  MoveL 5119 to (-200, -30.3, 0.2) mm, rotated rx 1.14 ry 0 rz 180 deg; joints [20.999, -64.73, 124.107, -155.961, 61.604, 79.168]
  MoveL 5120 to (0, -30.3, 0.2) mm, rotated rx 1.14 ry 0 rz 180 deg; joints [18.154, -55.53, 108.18, -157.586, 54.796, 77.769]
  MoveL 5121 to (0, -29.7, 0.2) mm, rotated rx 0 ry 0 rz 180 deg; joints [18.189, -55.157, 108.238, -157.658, 55.202, 76.801]
  MoveL 5122 to (-200, -29.7, 0.2) mm, rotated rx 0 ry 0 rz 180 deg; joints [21.039, -64.279, 124.171, -156.029, 62.083, 78.241]
  MoveL 5123 to (-200, -29.1, 0.2) mm, rotated rx 0 ry 0 rz 180 deg; joints [21.039, -64.245, 124.178, -156.038, 62.121, 78.259]
  MoveL 5124 to (0, -29.1, 0.2) mm, rotated rx 0 ry 0 rz 180 deg; joints [18.189, -55.13, 108.244, -157.667, 55.234, 76.816]
  MoveL 5125 to (0, -28.5, 0.2) mm, rotated rx 0 ry 0 rz 180 deg; joints [18.189, -55.102, 108.25, -157.676, 55.266, 76.832]
  MoveL 5126 to (-200, -28.5, 0.2) mm, rotated rx 0 ry 0 rz 180 deg; joints [21.039, -64.211, 124.185, -156.046, 62.158, 78.278]
  MoveL 5127 to (-200, -27.9, 0.2) mm, rotated rx 0 ry 0 rz 180 deg; joints [21.039, -64.177, 124.192, -156.055, 62.195, 78.297]
  MoveL 5128 to (0, -27.9, 0.2) mm, rotated rx 0 ry 0 rz 180 deg; joints [18.189, -55.074, 108.257, -157.685, 55.297, 76.848]
  MoveL 5129 to (0, -27.3, 0.2) mm, rotated rx 0 ry 0 rz 180 deg; joints [18.189, -55.046, 108.263, -157.694, 55.329, 76.864]
  MoveL 5130 to (-200, -27.3, 0.2) mm, rotated rx 0 ry 0 rz 180 deg; joints [21.039, -64.143, 124.198, -156.064, 62.232, 78.316]
  MoveL 5131 to (-200, -26.7, 0.2) mm, rotated rx 0 ry 0 rz 180 deg; joints [21.039, -64.109, 124.205, -156.072, 62.269, 78.334]
  MoveL 5132 to (0, -26.7, 0.2) mm, rotated rx 0 ry 0 rz 180 deg; joints [18.189, -55.018, 108.269, -157.703, 55.361, 76.88]
  MoveL 5133 to (0, -26.1, 0.2) mm, rotated rx 0 ry 0 rz 180 deg; joints [18.189, -54.99, 108.275, -157.712, 55.392, 76.895]
  MoveL 5134 to (-200, -26.1, 0.2) mm, rotated rx 0 ry 0 rz 180 deg; joints [21.039, -64.075, 124.212, -156.081, 62.307, 78.353]
  MoveL 5135 to (-200, -25.5, 0.2) mm, rotated rx 0 ry 0 rz 180 deg; joints [21.039, -64.041, 124.218, -156.09, 62.344, 78.372]
  MoveL 5136 to (0, -25.5, 0.2) mm, rotated rx 0 ry 0 rz 180 deg; joints [18.189, -54.962, 108.281, -157.721, 55.424, 76.911]
  MoveL 5137 to (0, -24.9, 0.2) mm, rotated rx 0 ry 0 rz 180 deg; joints [18.189, -54.934, 108.288, -157.73, 55.455, 76.927]
  MoveL 5138 to (-200, -24.9, 0.2) mm, rotated rx 0 ry 0 rz 180 deg; joints [21.039, -64.007, 124.225, -156.098, 62.381, 78.39]
  MoveL 5139 to (-200, -24.3, 0.2) mm, rotated rx 0 ry 0 rz 180 deg; joints [21.039, -63.973, 124.232, -156.107, 62.418, 78.409]
  MoveL 5140 to (0, -24.3, 0.2) mm, rotated rx 0 ry 0 rz 180 deg; joints [18.189, -54.906, 108.294, -157.739, 55.487, 76.942]
  MoveL 5141 to (0, -23.7, 0.2) mm, rotated rx 0 ry 0 rz 180 deg; joints [18.189, -54.878, 108.3, -157.748, 55.519, 76.958]
  MoveL 5142 to (-200, -23.7, 0.2) mm, rotated rx 0 ry 0 rz 180 deg; joints [21.039, -63.939, 124.238, -156.116, 62.455, 78.427]
  MoveL 5143 to (-200, -23.1, 0.2) mm, rotated rx 0 ry 0 rz 180 deg; joints [21.039, -63.905, 124.245, -156.124, 62.493, 78.446]
  MoveL 5144 to (0, -23.1, 0.2) mm, rotated rx 0 ry 0 rz 180 deg; joints [18.189, -54.849, 108.306, -157.757, 55.55, 76.974]
  MoveL 5145 to (0, -22.5, 0.2) mm, rotated rx 0 ry 0 rz 180 deg; joints [18.189, -54.821, 108.312, -157.766, 55.582, 76.989]
  MoveL 5146 to (-200, -22.5, 0.2) mm, rotated rx 0 ry 0 rz 180 deg; joints [21.039, -63.871, 124.251, -156.133, 62.53, 78.464]
  MoveL 5147 to (-200, -21.9, 0.2) mm, rotated rx 0 ry 0 rz 180 deg; joints [21.039, -63.836, 124.258, -156.141, 62.567, 78.483]
  MoveL 5148 to (0, -21.9, 0.2) mm, rotated rx 0 ry 0 rz 180 deg; joints [18.189, -54.793, 108.318, -157.775, 55.613, 77.005]
  MoveL 5149 to (0, -21.3, 0.2) mm, rotated rx 0 ry 0 rz 180 deg; joints [18.189, -54.765, 108.324, -157.783, 55.645, 77.021]
  MoveL 5150 to (-200, -21.3, 0.2) mm, rotated rx 0 ry 0 rz 180 deg; joints [21.039, -63.802, 124.264, -156.15, 62.604, 78.501]
  MoveL 5151 to (-200, -20.7, 0.2) mm, rotated rx 0 ry 0 rz 180 deg; joints [21.039, -63.768, 124.271, -156.158, 62.641, 78.52]
  MoveL 5152 to (0, -20.7, 0.2) mm, rotated rx 0 ry 0 rz 180 deg; joints [18.189, -54.737, 108.33, -157.792, 55.676, 77.036]
  MoveL 5153 to (0, -20.1, 0.2) mm, rotated rx 0 ry 0 rz 180 deg; joints [18.189, -54.709, 108.335, -157.801, 55.708, 77.052]
  MoveL 5154 to (-200, -20.1, 0.2) mm, rotated rx 0 ry 0 rz 180 deg; joints [21.039, -63.734, 124.277, -156.167, 62.678, 78.538]
  MoveL 5155 to (-200, -19.5, 0.2) mm, rotated rx 0 ry 0 rz 180 deg; joints [21.039, -63.7, 124.283, -156.175, 62.716, 78.557]
  MoveL 5156 to (0, -19.5, 0.2) mm, rotated rx 0 ry 0 rz 180 deg; joints [18.189, -54.681, 108.341, -157.81, 55.739, 77.067]
  MoveL 5157 to (0, -18.9, 0.2) mm, rotated rx 0 ry 0 rz 180 deg; joints [18.189, -54.652, 108.347, -157.818, 55.771, 77.083]
  MoveL 5158 to (-200, -18.9, 0.2) mm, rotated rx 0 ry 0 rz 180 deg; joints [21.039, -63.665, 124.29, -156.184, 62.753, 78.575]
  MoveL 5159 to (-200, -18.3, 0.2) mm, rotated rx 0 ry 0 rz 180 deg; joints [21.039, -63.631, 124.296, -156.192, 62.79, 78.594]
  MoveL 5160 to (0, -18.3, 0.2) mm, rotated rx 0 ry 0 rz 180 deg; joints [18.189, -54.624, 108.353, -157.827, 55.802, 77.099]
  MoveL 5161 to (0, -17.7, 0.2) mm, rotated rx 0 ry 0 rz 180 deg; joints [18.189, -54.596, 108.359, -157.836, 55.834, 77.114]
  MoveL 5162 to (-200, -17.7, 0.2) mm, rotated rx 0 ry 0 rz 180 deg; joints [21.039, -63.597, 124.302, -156.201, 62.827, 78.612]
  MoveL 5163 to (-200, -17.1, 0.2) mm, rotated rx 0 ry 0 rz 180 deg; joints [21.039, -63.562, 124.308, -156.209, 62.864, 78.631]
  MoveL 5164 to (0, -17.1, 0.2) mm, rotated rx 0 ry 0 rz 180 deg; joints [18.189, -54.568, 108.364, -157.845, 55.865, 77.13]
  MoveL 5165 to (0, -16.5, 0.2) mm, rotated rx 0 ry 0 rz 180 deg; joints [18.189, -54.539, 108.37, -157.853, 55.897, 77.145]
  MoveL 5166 to (-200, -16.5, 0.2) mm, rotated rx 0 ry 0 rz 180 deg; joints [21.039, -63.528, 124.315, -156.217, 62.901, 78.649]
  MoveL 5167 to (-200, -15.9, 0.2) mm, rotated rx 0 ry 0 rz 180 deg; joints [21.039, -63.494, 124.321, -156.226, 62.938, 78.667]
  MoveL 5168 to (0, -15.9, 0.2) mm, rotated rx 0 ry 0 rz 180 deg; joints [18.189, -54.511, 108.376, -157.862, 55.928, 77.161]
  MoveL 5169 to (0, -15.3, 0.2) mm, rotated rx 0 ry 0 rz 180 deg; joints [18.189, -54.483, 108.381, -157.871, 55.96, 77.176]
  MoveL 5170 to (-200, -15.3, 0.2) mm, rotated rx 0 ry 0 rz 180 deg; joints [21.039, -63.459, 124.327, -156.234, 62.975, 78.686]
  MoveL 5171 to (-200, -14.7, 0.2) mm, rotated rx 0 ry 0 rz 180 deg; joints [21.039, -63.425, 124.333, -156.242, 63.012, 78.704]
  MoveL 5172 to (0, -14.7, 0.2) mm, rotated rx 0 ry 0 rz 180 deg; joints [18.189, -54.454, 108.387, -157.879, 55.991, 77.191]
  MoveL 5173 to (0, -14.1, 0.2) mm, rotated rx 0 ry 0 rz 180 deg; joints [18.189, -54.426, 108.393, -157.888, 56.023, 77.207]
  MoveL 5174 to (-200, -14.1, 0.2) mm, rotated rx 0 ry 0 rz 180 deg; joints [21.039, -63.39, 124.339, -156.251, 63.049, 78.722]
  MoveL 5175 to (-200, -13.5, 0.2) mm, rotated rx 0 ry 0 rz 180 deg; joints [21.039, -63.356, 124.345, -156.259, 63.087, 78.741]
  MoveL 5176 to (0, -13.5, 0.2) mm, rotated rx 0 ry 0 rz 180 deg; joints [18.189, -54.398, 108.398, -157.896, 56.054, 77.222]
  MoveL 5177 to (0, -12.9, 0.2) mm, rotated rx 0 ry 0 rz 180 deg; joints [18.189, -54.369, 108.404, -157.905, 56.086, 77.238]
  MoveL 5178 to (-200, -12.9, 0.2) mm, rotated rx 0 ry 0 rz 180 deg; joints [21.039, -63.321, 124.351, -156.267, 63.124, 78.759]
  MoveL 5179 to (-200, -12.3, 0.2) mm, rotated rx 0 ry 0 rz 180 deg; joints [21.039, -63.287, 124.357, -156.275, 63.161, 78.777]
  MoveL 5180 to (0, -12.3, 0.2) mm, rotated rx 0 ry 0 rz 180 deg; joints [18.189, -54.341, 108.409, -157.914, 56.117, 77.253]
  MoveL 5181 to (0, -11.7, 0.2) mm, rotated rx 0 ry 0 rz 180 deg; joints [18.189, -54.312, 108.415, -157.922, 56.148, 77.268]
  MoveL 5182 to (-200, -11.7, 0.2) mm, rotated rx 0 ry 0 rz 180 deg; joints [21.039, -63.252, 124.363, -156.284, 63.198, 78.795]
  MoveL 5183 to (-200, -11.1, 0.2) mm, rotated rx 0 ry 0 rz 180 deg; joints [21.039, -63.218, 124.369, -156.292, 63.235, 78.814]
  MoveL 5184 to (0, -11.1, 0.2) mm, rotated rx 0 ry 0 rz 180 deg; joints [18.189, -54.284, 108.42, -157.931, 56.18, 77.284]
  MoveL 5185 to (0, -10.5, 0.2) mm, rotated rx 0 ry 0 rz 180 deg; joints [18.189, -54.256, 108.426, -157.939, 56.211, 77.299]
  MoveL 5186 to (-200, -10.5, 0.2) mm, rotated rx 0 ry 0 rz 180 deg; joints [21.039, -63.183, 124.375, -156.3, 63.272, 78.832]
  MoveL 5187 to (-200, -9.9, 0.2) mm, rotated rx 0 ry 0 rz 180 deg; joints [21.039, -63.149, 124.381, -156.308, 63.309, 78.85]
  MoveL 5188 to (0, -9.9, 0.2) mm, rotated rx 0 ry 0 rz 180 deg; joints [18.189, -54.227, 108.431, -157.948, 56.243, 77.314]
  MoveL 5189 to (0, -9.3, 0.2) mm, rotated rx 0 ry 0 rz 180 deg; joints [18.189, -54.199, 108.436, -157.956, 56.274, 77.33]
  MoveL 5190 to (-200, -9.3, 0.2) mm, rotated rx 0 ry 0 rz 180 deg; joints [21.039, -63.114, 124.387, -156.316, 63.346, 78.868]
  MoveL 5191 to (-200, -8.7, 0.2) mm, rotated rx 0 ry 0 rz 180 deg; joints [21.039, -63.079, 124.392, -156.325, 63.383, 78.886]
  MoveL 5192 to (0, -8.7, 0.2) mm, rotated rx 0 ry 0 rz 180 deg; joints [18.189, -54.17, 108.442, -157.965, 56.305, 77.345]
  MoveL 5193 to (0, -8.1, 0.2) mm, rotated rx 0 ry 0 rz 180 deg; joints [18.189, -54.141, 108.447, -157.973, 56.337, 77.36]
  MoveL 5194 to (-200, -8.1, 0.2) mm, rotated rx 0 ry 0 rz 180 deg; joints [21.039, -63.045, 124.398, -156.333, 63.42, 78.904]
  MoveL 5195 to (-200, -7.5, 0.2) mm, rotated rx 0 ry 0 rz 180 deg; joints [21.039, -63.01, 124.404, -156.341, 63.457, 78.923]
  MoveL 5196 to (0, -7.5, 0.2) mm, rotated rx 0 ry 0 rz 180 deg; joints [18.189, -54.113, 108.452, -157.982, 56.368, 77.375]
  MoveL 5197 to (0, -6.9, 0.2) mm, rotated rx 0 ry 0 rz 180 deg; joints [18.189, -54.084, 108.457, -157.99, 56.399, 77.391]
  MoveL 5198 to (-200, -6.9, 0.2) mm, rotated rx 0 ry 0 rz 180 deg; joints [21.039, -62.975, 124.409, -156.349, 63.494, 78.941]
  MoveL 5199 to (-200, -6.3, 0.2) mm, rotated rx 0 ry 0 rz 180 deg; joints [21.039, -62.941, 124.415, -156.357, 63.531, 78.959]
  MoveL 5200 to (0, -6.3, 0.2) mm, rotated rx 0 ry 0 rz 180 deg; joints [18.189, -54.056, 108.463, -157.998, 56.431, 77.406]
  MoveL 5201 to (0, -5.7, 0.2) mm, rotated rx 0 ry 0 rz 180 deg; joints [18.189, -54.027, 108.468, -158.007, 56.462, 77.421]
  MoveL 5202 to (-200, -5.7, 0.2) mm, rotated rx 0 ry 0 rz 180 deg; joints [21.039, -62.906, 124.421, -156.365, 63.568, 78.977]
  MoveL 5203 to (-200, -5.1, 0.2) mm, rotated rx 0 ry 0 rz 180 deg; joints [21.039, -62.871, 124.426, -156.373, 63.605, 78.995]
  MoveL 5204 to (0, -5.1, 0.2) mm, rotated rx 0 ry 0 rz 180 deg; joints [18.189, -53.999, 108.473, -158.015, 56.493, 77.436]
  MoveL 5205 to (0, -4.5, 0.2) mm, rotated rx 0 ry 0 rz 180 deg; joints [18.189, -53.97, 108.478, -158.024, 56.525, 77.451]
  MoveL 5206 to (-200, -4.5, 0.2) mm, rotated rx 0 ry 0 rz 180 deg; joints [21.039, -62.836, 124.432, -156.381, 63.642, 79.013]
  MoveL 5207 to (-200, -3.9, 0.2) mm, rotated rx 0 ry 0 rz 180 deg; joints [21.039, -62.802, 124.437, -156.389, 63.679, 79.031]
  MoveL 5208 to (0, -3.9, 0.2) mm, rotated rx 0 ry 0 rz 180 deg; joints [18.189, -53.941, 108.483, -158.032, 56.556, 77.466]
  MoveL 5209 to (0, -3.3, 0.2) mm, rotated rx 0 ry 0 rz 180 deg; joints [18.189, -53.913, 108.488, -158.04, 56.587, 77.481]
  MoveL 5210 to (-200, -3.3, 0.2) mm, rotated rx 0 ry 0 rz 180 deg; joints [21.039, -62.767, 124.443, -156.397, 63.716, 79.049]
  MoveL 5211 to (-200, -2.7, 0.2) mm, rotated rx 0 ry 0 rz 180 deg; joints [21.039, -62.732, 124.448, -156.405, 63.753, 79.067]
  MoveL 5212 to (0, -2.7, 0.2) mm, rotated rx 0 ry 0 rz 180 deg; joints [18.189, -53.884, 108.493, -158.049, 56.619, 77.497]
  MoveL 5213 to (0, -2.1, 0.2) mm, rotated rx 0 ry 0 rz 180 deg; joints [18.189, -53.855, 108.498, -158.057, 56.65, 77.512]
  MoveL 5214 to (-200, -2.1, 0.2) mm, rotated rx 0 ry 0 rz 180 deg; joints [21.039, -62.697, 124.454, -156.413, 63.789, 79.085]
  MoveL 5215 to (-200, -1.5, 0.2) mm, rotated rx 0 ry 0 rz 180 deg; joints [21.039, -62.662, 124.459, -156.421, 63.826, 79.103]
  MoveL 5216 to (0, -1.5, 0.2) mm, rotated rx 0 ry 0 rz 180 deg; joints [18.189, -53.826, 108.503, -158.065, 56.681, 77.527]
  MoveL 5217 to (0, -0.9, 0.2) mm, rotated rx 0 ry 0 rz 180 deg; joints [18.189, -53.798, 108.508, -158.073, 56.712, 77.542]
  MoveL 5218 to (-200, -0.9, 0.2) mm, rotated rx 0 ry 0 rz 180 deg; joints [21.039, -62.627, 124.465, -156.429, 63.863, 79.121]
  MoveL 5219 to (-200, -0.3, 0.2) mm, rotated rx 0 ry 0 rz 180 deg; joints [21.039, -62.592, 124.47, -156.437, 63.9, 79.139]
  MoveL 5220 to (0, -0.3, 0.2) mm, rotated rx 0 ry 0 rz 180 deg; joints [18.189, -53.769, 108.513, -158.082, 56.744, 77.557]
  MoveL 5221 to (0, 0, 0.2) mm, rotated rx 0 ry 0 rz 180 deg; joints [18.189, -53.755, 108.515, -158.086, 56.759, 77.564]
  MoveL 5222 to (-200, 0, 0.2) mm, rotated rx 0 ry 0 rz 180 deg; joints [21.039, -62.575, 124.473, -156.44, 63.918, 79.148]
  Sollgeschwindigkeit (200.0 mm/s)
  MoveL 5223 to (-200, 0, -44.8) mm, rotated rx 0 ry 0 rz 180 deg; joints [22.93, -61.804, 123.11, -154.254, 63.757, 77.962]
  END

--- program CBL1 (robot KUKA KR 30 HA) ---
  Glatt(1)
  Sollgeschwindigkeit (1000.0 mm/s)
  Referenz erstellen.: Reference SW
  Werkzeug setzen: PlasticPos800
  Anzeigen PlasticPos800
  MoveJ 1 to (-41.72, -40.46, 48.98) mm, rotated rx 90 ry 0 rz 90 deg; joints [0.027, -82.593, 139.4, -179.968, 56.807, 179.983]
  MoveL 2 to (-41.72, -40.46, 48.98) mm, rotated rx 90 ry 0 rz 90 deg; joints [0.027, -82.593, 139.4, -179.968, 56.807, 179.983]
  MoveL 3 to (-41.72, -40.46, 48.98) mm, rotated rx 90 ry 0 rz 90 deg; joints [0.027, -82.593, 139.4, -179.968, 56.807, 179.983]
  MoveL 4 to (-41.72, -40.46, 48.98) mm, rotated rx 90 ry 0 rz 90 deg; joints [0.027, -82.593, 139.4, -179.968, 56.807, 179.983]
  Sollgeschwindigkeit (50.0 mm/s)
  MoveL 5 to (-32.85, -40.57, 48.4) mm, rotated rx 90 ry 0 rz 90 deg; joints [0.058, -82.072, 138.764, -179.93, 56.692, 179.962]
  MoveL 6 to (-23.97, -40.69, 47.75) mm, rotated rx 90 ry 0 rz 90 deg; joints [0.094, -81.555, 138.126, -179.887, 56.571, 179.938]
  MoveL 7 to (-15.09, -40.74, 47.81) mm, rotated rx 90 ry 0 rz 90 deg; joints [0.089, -81.036, 137.485, -179.893, 56.449, 179.941]
  MoveL 8 to (-6.28, -40.47, 49.1) mm, rotated rx 90 ry 0 rz 90 deg; joints [0.02, -80.506, 136.856, -179.976, 56.35, 179.987]
  MoveL 9 to (-0.84, -39.84, 50.5) mm, rotated rx 90 ry 0 rz 90 deg; joints [-0.055, -80.152, 136.477, -180.066, 56.326, 180.037]
  MoveL 10 to (4.48, -38.76, 52.1) mm, rotated rx 90 ry 0 rz 90 deg; joints [-0.14, -79.779, 136.116, -180.168, 56.337, 180.093]
  MoveL 11 to (9.75, -37.21, 53.58) mm, rotated rx 90 ry 0 rz 90 deg; joints [-0.218, -79.383, 135.768, -180.262, 56.385, 180.145]
  MoveL 12 to (14.99, -35.35, 54.76) mm, rotated rx 90 ry 0 rz 90 deg; joints [-0.279, -78.971, 135.428, -180.335, 56.457, 180.185]
  MoveL 13 to (20.23, -33.45, 55.56) mm, rotated rx 90 ry 0 rz 90 deg; joints [-0.32, -78.559, 135.087, -180.383, 56.528, 180.212]
  MoveL 14 to (25.53, -31.86, 55.96) mm, rotated rx 90 ry 0 rz 90 deg; joints [-0.339, -78.165, 134.733, -180.407, 56.569, 180.224]
  MoveL 15 to (31.11, -31.04, 56.06) mm, rotated rx 90 ry 0 rz 90 deg; joints [-0.343, -77.802, 134.34, -180.411, 56.539, 180.227]
  MoveL 16 to (37.22, -31.47, 56) mm, rotated rx 90 ry 0 rz 90 deg; joints [-0.338, -77.485, 133.88, -180.405, 56.395, 180.224]
  MoveL 17 to (43.65, -32.9, 55.86) mm, rotated rx 90 ry 0 rz 90 deg; joints [-0.329, -77.209, 133.372, -180.396, 56.164, 180.22]
  MoveL 18 to (50.35, -33.59, 55.79) mm, rotated rx 90 ry 0 rz 90 deg; joints [-0.323, -76.875, 132.859, -180.39, 55.985, 180.218]
  MoveL 19 to (57.02, -32.75, 55.87) mm, rotated rx 90 ry 0 rz 90 deg; joints [-0.325, -76.455, 132.381, -180.393, 55.926, 180.22]
  MoveL 20 to (63.44, -31.36, 56.01) mm, rotated rx 90 ry 0 rz 90 deg; joints [-0.33, -76.02, 131.931, -180.399, 55.912, 180.224]
  MoveL 21 to (69.49, -31.08, 56.06) mm, rotated rx 90 ry 0 rz 90 deg; joints [-0.331, -75.67, 131.484, -180.401, 55.815, 180.225]
  MoveL 22 to (75.02, -32, 55.94) mm, rotated rx 90 ry 0 rz 90 deg; joints [-0.323, -75.417, 131.048, -180.392, 55.631, 180.221]
  MoveL 23 to (80.31, -33.64, 55.49) mm, rotated rx 90 ry 0 rz 90 deg; joints [-0.3, -75.218, 130.615, -180.364, 55.397, 180.207]
  MoveL 24 to (85.55, -35.55, 54.65) mm, rotated rx 90 ry 0 rz 90 deg; joints [-0.257, -75.036, 130.178, -180.313, 55.143, 180.179]
  MoveL 25 to (93.19, -38.13, 52.78) mm, rotated rx 90 ry 0 rz 90 deg; joints [-0.163, -74.758, 129.545, -180.2, 54.787, 180.115]
  MoveL 26 to (100.91, -39.85, 50.48) mm, rotated rx 90 ry 0 rz 90 deg; joints [-0.049, -74.427, 128.922, -180.061, 54.495, 180.035]
  MoveL 27 to (108.88, -40.62, 48.59) mm, rotated rx 90 ry 0 rz 90 deg; joints [0.042, -74.031, 128.298, -179.948, 54.266, 179.969]
  MoveL 28 to (117.07, -40.74, 47.7) mm, rotated rx 90 ry 0 rz 90 deg; joints [0.085, -73.589, 127.669, -179.895, 54.08, 179.938]
  MoveL 29 to (125.29, -40.67, 47.82) mm, rotated rx 90 ry 0 rz 90 deg; joints [0.079, -73.136, 127.039, -179.903, 53.902, 179.943]
  MoveL 30 to (133.51, -40.57, 48.46) mm, rotated rx 90 ry 0 rz 90 deg; joints [0.048, -72.683, 126.408, -179.941, 53.724, 179.965]
  MoveL 31 to (141.72, -40.46, 48.98) mm, rotated rx 90 ry 0 rz 90 deg; joints [0.023, -72.231, 125.774, -179.972, 53.543, 179.983]
  Sollgeschwindigkeit (1000.0 mm/s)
  MoveL 32 to (141.72, -40.46, 48.98) mm, rotated rx 90 ry 0 rz 90 deg; joints [0.023, -72.231, 125.774, -179.972, 53.543, 179.983]
  MoveL 33 to (141.72, -40.46, 48.98) mm, rotated rx 90 ry 0 rz 90 deg; joints [0.023, -72.231, 125.774, -179.972, 53.543, 179.983]
  Sollgeschwindigkeit (1000.0 mm/s)
  MoveL 34 to (145.1, -41.25, 44.7) mm, rotated rx 90 ry 0 rz 90 deg; joints [0.224, -72.088, 125.494, -179.721, 53.406, 179.834]
  MoveL 35 to (145.1, -41.25, 44.7) mm, rotated rx 90 ry 0 rz 90 deg; joints [0.224, -72.088, 125.494, -179.721, 53.406, 179.834]
  MoveL 36 to (145.1, -41.25, 44.7) mm, rotated rx 90 ry 0 rz 90 deg; joints [0.224, -72.088, 125.494, -179.721, 53.406, 179.834]
  Sollgeschwindigkeit (50.0 mm/s)
  MoveL 37 to (141.7, -41.25, 42.87) mm, rotated rx 90 ry 0 rz 90 deg; joints [0.312, -72.273, 125.758, -179.612, 53.486, 179.769]
  MoveL 38 to (137.92, -41.25, 41.96) mm, rotated rx 90 ry 0 rz 90 deg; joints [0.355, -72.478, 126.05, -179.558, 53.573, 179.738]
  MoveL 39 to (134, -41.25, 41.48) mm, rotated rx 90 ry 0 rz 90 deg; joints [0.379, -72.691, 126.353, -179.529, 53.663, 179.721]
  MoveL 40 to (130.09, -41.25, 41.08) mm, rotated rx 90 ry 0 rz 90 deg; joints [0.4, -72.903, 126.655, -179.505, 53.752, 179.707]
  MoveL 41 to (126.21, -41.24, 40.71) mm, rotated rx 90 ry 0 rz 90 deg; joints [0.419, -73.115, 126.954, -179.481, 53.84, 179.694]
  MoveL 42 to (118.64, -41.24, 39.88) mm, rotated rx 90 ry 0 rz 90 deg; joints [0.461, -73.528, 127.535, -179.43, 54.008, 179.665]
  MoveL 43 to (111.13, -41.25, 38.67) mm, rotated rx 90 ry 0 rz 90 deg; joints [0.523, -73.939, 128.109, -179.355, 54.171, 179.623]
  MoveL 44 to (104.5, -41.27, 37.04) mm, rotated rx 90 ry 0 rz 90 deg; joints [0.605, -74.303, 128.613, -179.255, 54.312, 179.565]
  MoveL 45 to (98.04, -41.26, 34.74) mm, rotated rx 90 ry 0 rz 90 deg; joints [0.721, -74.656, 129.102, -179.113, 54.449, 179.485]
  MoveL 46 to (91.88, -41.2, 31.62) mm, rotated rx 90 ry 0 rz 90 deg; joints [0.879, -74.99, 129.567, -178.922, 54.581, 179.375]
  MoveL 47 to (86.28, -41.2, 27.66) mm, rotated rx 90 ry 0 rz 90 deg; joints [1.079, -75.296, 129.985, -178.678, 54.697, 179.236]
  MoveL 48 to (80.96, -41.38, 22.17) mm, rotated rx 90 ry 0 rz 90 deg; joints [1.356, -75.594, 130.373, -178.34, 54.791, 179.043]
  MoveL 49 to (76.3, -41.22, 15.86) mm, rotated rx 90 ry 0 rz 90 deg; joints [1.677, -75.835, 130.715, -177.95, 54.897, 178.821]
  MoveL 50 to (73.92, -40.67, 12.58) mm, rotated rx 90 ry 0 rz 90 deg; joints [1.844, -75.931, 130.898, -177.748, 54.988, 178.708]
  MoveL 51 to (71.58, -39.57, 9.53) mm, rotated rx 90 ry 0 rz 90 deg; joints [2.001, -75.994, 131.09, -177.561, 55.121, 178.605]
  MoveL 52 to (69.42, -37.75, 7.01) mm, rotated rx 90 ry 0 rz 90 deg; joints [2.131, -76.007, 131.286, -177.408, 55.306, 178.524]
  MoveL 53 to (67.55, -35.05, 5.3) mm, rotated rx 90 ry 0 rz 90 deg; joints [2.22, -75.955, 131.48, -177.307, 55.555, 178.476]
  MoveL 54 to (65.46, -30.42, 4.14) mm, rotated rx 90 ry 0 rz 90 deg; joints [2.283, -75.806, 131.734, -177.245, 55.959, 178.457]
  MoveL 55 to (63.59, -25.34, 3.78) mm, rotated rx 90 ry 0 rz 90 deg; joints [2.305, -75.618, 131.981, -177.233, 56.394, 178.468]
  MoveL 56 to (61.65, -20.55, 3.71) mm, rotated rx 90 ry 0 rz 90 deg; joints [2.312, -75.447, 132.227, -177.237, 56.81, 178.487]
  MoveL 57 to (59.77, -17.22, 3.72) mm, rotated rx 90 ry 0 rz 90 deg; joints [2.315, -75.355, 132.436, -177.243, 57.111, 178.502]
  MoveL 58 to (57.13, -13.98, 3.77) mm, rotated rx 90 ry 0 rz 90 deg; joints [2.318, -75.309, 132.7, -177.248, 57.421, 178.518]
  MoveL 59 to (55.51, -12.44, 3.79) mm, rotated rx 90 ry 0 rz 90 deg; joints [2.32, -75.305, 132.851, -177.251, 57.576, 178.525]
  MoveL 60 to (53.83, -11.08, 3.81) mm, rotated rx 90 ry 0 rz 90 deg; joints [2.323, -75.316, 133.004, -177.252, 57.718, 178.531]
  MoveL 61 to (52.14, -9.99, 3.81) mm, rotated rx 90 ry 0 rz 90 deg; joints [2.327, -75.342, 133.153, -177.251, 57.84, 178.536]
  MoveL 62 to (50, -9.51, 3.8) mm, rotated rx 90 ry 0 rz 90 deg; joints [2.331, -75.43, 133.322, -177.248, 57.923, 178.538]
  MoveL 63 to (47.86, -9.99, 3.81) mm, rotated rx 90 ry 0 rz 90 deg; joints [2.336, -75.574, 133.473, -177.243, 57.929, 178.536]
  MoveL 64 to (46.17, -11.08, 3.81) mm, rotated rx 90 ry 0 rz 90 deg; joints [2.339, -75.731, 133.577, -177.238, 57.876, 178.53]
  MoveL 65 to (44.49, -12.44, 3.79) mm, rotated rx 90 ry 0 rz 90 deg; joints [2.343, -75.904, 133.675, -177.23, 57.801, 178.523]
  MoveL 66 to (42.87, -13.98, 3.77) mm, rotated rx 90 ry 0 rz 90 deg; joints [2.348, -76.084, 133.764, -177.222, 57.711, 178.515]
  MoveL 67 to (40.23, -17.22, 3.72) mm, rotated rx 90 ry 0 rz 90 deg; joints [2.356, -76.422, 133.894, -177.207, 57.503, 178.498]
  MoveL 68 to (38.35, -20.55, 3.71) mm, rotated rx 90 ry 0 rz 90 deg; joints [2.36, -76.725, 133.963, -177.194, 57.27, 178.482]
  MoveL 69 to (36.41, -25.34, 3.78) mm, rotated rx 90 ry 0 rz 90 deg; joints [2.361, -77.117, 134.005, -177.182, 56.92, 178.461]
  MoveL 70 to (34.54, -30.42, 4.14) mm, rotated rx 90 ry 0 rz 90 deg; joints [2.346, -77.522, 134.034, -177.187, 56.543, 178.448]
  MoveL 71 to (32.45, -35.05, 5.3) mm, rotated rx 90 ry 0 rz 90 deg; joints [2.291, -77.915, 134.089, -177.243, 56.205, 178.466]
  MoveL 72 to (30.58, -37.75, 7.01) mm, rotated rx 90 ry 0 rz 90 deg; joints [2.206, -78.182, 134.17, -177.339, 56.016, 178.512]
  MoveL 73 to (28.42, -39.57, 9.53) mm, rotated rx 90 ry 0 rz 90 deg; joints [2.079, -78.417, 134.294, -177.489, 55.902, 178.592]
  MoveL 74 to (26.08, -40.67, 12.58) mm, rotated rx 90 ry 0 rz 90 deg; joints [1.925, -78.62, 134.448, -177.674, 55.85, 178.694]
  MoveL 75 to (23.7, -41.22, 15.86) mm, rotated rx 90 ry 0 rz 90 deg; joints [1.757, -78.794, 134.617, -177.876, 55.841, 178.807]
  MoveL 76 to (19.04, -41.38, 22.17) mm, rotated rx 90 ry 0 rz 90 deg; joints [1.433, -79.079, 134.968, -178.269, 55.9, 179.029]
  MoveL 77 to (13.72, -41.2, 27.66) mm, rotated rx 90 ry 0 rz 90 deg; joints [1.151, -79.381, 135.37, -178.612, 55.997, 179.224]
  MoveL 78 to (6.48, -41.22, 32.56) mm, rotated rx 90 ry 0 rz 90 deg; joints [0.899, -79.804, 135.903, -178.918, 56.104, 179.396]
  MoveL 79 to (-1.54, -41.27, 36.09) mm, rotated rx 90 ry 0 rz 90 deg; joints [0.716, -80.274, 136.488, -179.138, 56.217, 179.521]
  MoveL 80 to (-9.91, -41.26, 38.42) mm, rotated rx 90 ry 0 rz 90 deg; joints [0.596, -80.762, 137.096, -179.284, 56.336, 179.603]
  MoveL 81 to (-18.44, -41.24, 39.85) mm, rotated rx 90 ry 0 rz 90 deg; joints [0.523, -81.261, 137.711, -179.373, 56.452, 179.653]
  MoveL 82 to (-33.66, -41.25, 41.44) mm, rotated rx 90 ry 0 rz 90 deg; joints [0.443, -82.161, 138.803, -179.47, 56.643, 179.709]
  MoveL 83 to (-37.69, -41.25, 41.93) mm, rotated rx 90 ry 0 rz 90 deg; joints [0.418, -82.401, 139.091, -179.5, 56.691, 179.726]
  MoveL 84 to (-41.59, -41.25, 42.83) mm, rotated rx 90 ry 0 rz 90 deg; joints [0.369, -82.634, 139.369, -179.559, 56.736, 179.758]
  MoveL 85 to (-45.1, -41.25, 44.7) mm, rotated rx 90 ry 0 rz 90 deg; joints [0.266, -82.845, 139.62, -179.682, 56.775, 179.826]
  Sollgeschwindigkeit (1000.0 mm/s)
  MoveL 86 to (-45.1, -41.25, 44.7) mm, rotated rx 90 ry 0 rz 90 deg; joints [0.266, -82.845, 139.62, -179.682, 56.775, 179.826]
  MoveL 87 to (-45.1, -41.25, 44.7) mm, rotated rx 90 ry 0 rz 90 deg; joints [0.266, -82.845, 139.62, -179.682, 56.775, 179.826]
  Sollgeschwindigkeit (1000.0 mm/s)
  MoveL 88 to (-50, -41.25, 39.09) mm, rotated rx 90 ry 0 rz 90 deg; joints [0.582, -83.137, 139.964, -179.305, 56.83, 179.62]
  MoveL 89 to (-50, -41.25, 39.09) mm, rotated rx 90 ry 0 rz 90 deg; joints [0.582, -83.137, 139.964, -179.305, 56.83, 179.62]
  MoveL 90 to (-50, -41.25, 39.09) mm, rotated rx 90 ry 0 rz 90 deg; joints [0.582, -83.137, 139.964, -179.305, 56.83, 179.62]
  Sollgeschwindigkeit (50.0 mm/s)
  MoveL 91 to (-43.32, -41.25, 37.37) mm, rotated rx 90 ry 0 rz 90 deg; joints [0.674, -82.734, 139.489, -179.195, 56.757, 179.558]
  MoveL 92 to (-36.74, -41.25, 35.17) mm, rotated rx 90 ry 0 rz 90 deg; joints [0.791, -82.34, 139.018, -179.053, 56.682, 179.48]
  MoveL 93 to (-30.13, -41.25, 33.25) mm, rotated rx 90 ry 0 rz 90 deg; joints [0.892, -81.946, 138.544, -178.932, 56.603, 179.412]
  MoveL 94 to (-23.34, -41.26, 32.21) mm, rotated rx 90 ry 0 rz 90 deg; joints [0.943, -81.545, 138.056, -178.87, 56.516, 179.376]
  MoveL 95 to (-16.33, -41.26, 31.5) mm, rotated rx 90 ry 0 rz 90 deg; joints [0.975, -81.132, 137.552, -178.829, 56.425, 179.353]
  MoveL 96 to (-9.37, -41.2, 30.15) mm, rotated rx 90 ry 0 rz 90 deg; joints [1.042, -80.72, 137.049, -178.748, 56.336, 179.306]
  MoveL 97 to (-2.68, -41.17, 27.82) mm, rotated rx 90 ry 0 rz 90 deg; joints [1.16, -80.327, 136.563, -178.605, 56.245, 179.225]
  MoveL 98 to (3.46, -41.31, 24.48) mm, rotated rx 90 ry 0 rz 90 deg; joints [1.331, -79.976, 136.109, -178.397, 56.144, 179.107]
  MoveL 99 to (8.93, -41.53, 20.18) mm, rotated rx 90 ry 0 rz 90 deg; joints [1.553, -79.666, 135.698, -178.128, 56.046, 178.954]
  MoveL 100 to (11.76, -41.47, 17.39) mm, rotated rx 90 ry 0 rz 90 deg; joints [1.696, -79.496, 135.488, -177.955, 56.009, 178.856]
  MoveL 101 to (14.45, -41.15, 14.37) mm, rotated rx 90 ry 0 rz 90 deg; joints [1.851, -79.316, 135.292, -177.767, 55.996, 178.751]
  MoveL 102 to (17.02, -40.42, 11.23) mm, rotated rx 90 ry 0 rz 90 deg; joints [2.012, -79.12, 135.114, -177.574, 56.018, 178.643]
  MoveL 103 to (19.34, -39.05, 8.37) mm, rotated rx 90 ry 0 rz 90 deg; joints [2.157, -78.9, 134.968, -177.4, 56.096, 178.549]
  MoveL 104 to (21.32, -36.78, 6.19) mm, rotated rx 90 ry 0 rz 90 deg; joints [2.268, -78.648, 134.87, -177.273, 56.251, 178.484]
  MoveL 105 to (22.97, -33.63, 4.84) mm, rotated rx 90 ry 0 rz 90 deg; joints [2.335, -78.365, 134.816, -177.199, 56.483, 178.453]
  MoveL 106 to (24.46, -29.95, 4.12) mm, rotated rx 90 ry 0 rz 90 deg; joints [2.369, -78.059, 134.787, -177.167, 56.76, 178.446]
  MoveL 107 to (26.01, -26.09, 3.8) mm, rotated rx 90 ry 0 rz 90 deg; joints [2.382, -77.742, 134.757, -177.16, 57.048, 178.455]
  MoveL 108 to (29.8, -19.01, 3.63) mm, rotated rx 90 ry 0 rz 90 deg; joints [2.383, -77.104, 134.629, -177.176, 57.556, 178.484]
  MoveL 109 to (34.48, -12.81, 3.73) mm, rotated rx 90 ry 0 rz 90 deg; joints [2.368, -76.472, 134.412, -177.207, 57.97, 178.518]
  MoveL 110 to (39.73, -7.1, 3.87) mm, rotated rx 90 ry 0 rz 90 deg; joints [2.35, -75.84, 134.136, -177.239, 58.326, 178.549]
  MoveL 111 to (45.25, -1.48, 3.82) mm, rotated rx 90 ry 0 rz 90 deg; joints [2.34, -75.201, 133.834, -177.26, 58.663, 178.574]
  Sollgeschwindigkeit (1000.0 mm/s)
  MoveL 112 to (45.25, -1.48, 3.82) mm, rotated rx 90 ry 0 rz 90 deg; joints [2.34, -75.201, 133.834, -177.26, 58.663, 178.574]
  MoveL 113 to (45.25, -1.48, 3.82) mm, rotated rx 90 ry 0 rz 90 deg; joints [2.34, -75.201, 133.834, -177.26, 58.663, 178.574]
  Sollgeschwindigkeit (1000.0 mm/s)
  MoveL 114 to (54.75, -1.48, 3.82) mm, rotated rx 90 ry 0 rz 90 deg; joints [2.321, -74.693, 133.123, -177.277, 58.459, 178.575]
  MoveL 115 to (54.75, -1.48, 3.82) mm, rotated rx 90 ry 0 rz 90 deg; joints [2.321, -74.693, 133.123, -177.277, 58.459, 178.575]
  MoveL 116 to (54.75, -1.48, 3.82) mm, rotated rx 90 ry 0 rz 90 deg; joints [2.321, -74.693, 133.123, -177.277, 58.459, 178.575]
  Sollgeschwindigkeit (50.0 mm/s)
  MoveL 117 to (60.27, -7.1, 3.87) mm, rotated rx 90 ry 0 rz 90 deg; joints [2.307, -74.733, 132.601, -177.276, 57.897, 178.552]
  MoveL 118 to (65.52, -12.81, 3.73) mm, rotated rx 90 ry 0 rz 90 deg; joints [2.303, -74.786, 132.093, -177.264, 57.336, 178.522]
  MoveL 119 to (70.2, -19.01, 3.63) mm, rotated rx 90 ry 0 rz 90 deg; joints [2.299, -74.893, 131.615, -177.251, 56.753, 178.492]
  MoveL 120 to (73.99, -26.09, 3.8) mm, rotated rx 90 ry 0 rz 90 deg; joints [2.283, -75.092, 131.184, -177.25, 56.123, 178.466]
  MoveL 121 to (75.54, -29.95, 4.12) mm, rotated rx 90 ry 0 rz 90 deg; joints [2.264, -75.226, 130.988, -177.262, 55.792, 178.46]
  MoveL 122 to (77.03, -33.63, 4.84) mm, rotated rx 90 ry 0 rz 90 deg; joints [2.225, -75.352, 130.798, -177.299, 55.476, 178.469]
  MoveL 123 to (78.68, -36.78, 6.19) mm, rotated rx 90 ry 0 rz 90 deg; joints [2.155, -75.439, 130.609, -177.376, 55.199, 178.502]
  MoveL 124 to (80.66, -39.05, 8.37) mm, rotated rx 90 ry 0 rz 90 deg; joints [2.043, -75.46, 130.417, -177.506, 54.983, 178.568]
  MoveL 125 to (82.98, -40.42, 11.23) mm, rotated rx 90 ry 0 rz 90 deg; joints [1.897, -75.412, 130.219, -177.68, 54.829, 178.663]
  MoveL 126 to (85.55, -41.15, 14.37) mm, rotated rx 90 ry 0 rz 90 deg; joints [1.737, -75.316, 130.017, -177.872, 54.72, 178.77]
  MoveL 127 to (88.24, -41.47, 17.39) mm, rotated rx 90 ry 0 rz 90 deg; joints [1.584, -75.189, 129.813, -178.058, 54.639, 178.876]
  MoveL 128 to (91.07, -41.53, 20.18) mm, rotated rx 90 ry 0 rz 90 deg; joints [1.443, -75.04, 129.604, -178.229, 54.576, 178.973]
  MoveL 129 to (96.54, -41.31, 24.48) mm, rotated rx 90 ry 0 rz 90 deg; joints [1.225, -74.732, 129.201, -178.495, 54.478, 179.125]
  MoveL 130 to (102.68, -41.17, 27.82) mm, rotated rx 90 ry 0 rz 90 deg; joints [1.056, -74.39, 128.743, -178.701, 54.36, 179.243]
  MoveL 131 to (109.37, -41.2, 30.15) mm, rotated rx 90 ry 0 rz 90 deg; joints [0.937, -74.027, 128.236, -178.845, 54.215, 179.325]
  MoveL 132 to (116.33, -41.26, 31.5) mm, rotated rx 90 ry 0 rz 90 deg; joints [0.866, -73.649, 127.704, -178.93, 54.059, 179.372]
  MoveL 133 to (123.34, -41.26, 32.21) mm, rotated rx 90 ry 0 rz 90 deg; joints [0.827, -73.267, 127.166, -178.976, 53.904, 179.397]
  MoveL 134 to (130.13, -41.25, 33.25) mm, rotated rx 90 ry 0 rz 90 deg; joints [0.773, -72.897, 126.646, -179.042, 53.753, 179.433]
  MoveL 135 to (136.74, -41.25, 35.17) mm, rotated rx 90 ry 0 rz 90 deg; joints [0.678, -72.538, 126.137, -179.158, 53.601, 179.5]
  MoveL 136 to (143.32, -41.25, 37.37) mm, rotated rx 90 ry 0 rz 90 deg; joints [0.57, -72.182, 125.629, -179.29, 53.449, 179.577]
  MoveL 137 to (150, -41.25, 39.09) mm, rotated rx 90 ry 0 rz 90 deg; joints [0.487, -71.821, 125.11, -179.393, 53.291, 179.637]
  Sollgeschwindigkeit (1000.0 mm/s)
  MoveL 138 to (150, -41.25, 39.09) mm, rotated rx 90 ry 0 rz 90 deg; joints [0.487, -71.821, 125.11, -179.393, 53.291, 179.637]
  MoveL 139 to (150, -41.25, 39.09) mm, rotated rx 90 ry 0 rz 90 deg; joints [0.487, -71.821, 125.11, -179.393, 53.291, 179.637]
  Sollgeschwindigkeit (1000.0 mm/s)
  MoveL 140 to (150, -41.25, 31.96) mm, rotated rx 90 ry 0 rz 90 deg; joints [0.821, -71.816, 125.104, -178.976, 53.292, 179.388]
  MoveL 141 to (150, -41.25, 31.96) mm, rotated rx 90 ry 0 rz 90 deg; joints [0.821, -71.816, 125.104, -178.976, 53.292, 179.388]
  MoveL 142 to (150, -41.25, 31.96) mm, rotated rx 90 ry 0 rz 90 deg; joints [0.821, -71.816, 125.104, -178.976, 53.292, 179.388]
  Sollgeschwindigkeit (50.0 mm/s)
  MoveL 143 to (144.93, -41.25, 28.57) mm, rotated rx 90 ry 0 rz 90 deg; joints [0.984, -72.088, 125.494, -178.774, 53.412, 179.269]
  MoveL 144 to (139.36, -41.27, 26.34) mm, rotated rx 90 ry 0 rz 90 deg; joints [1.094, -72.39, 125.923, -178.64, 53.541, 179.192]
  MoveL 145 to (133.44, -41.28, 24.88) mm, rotated rx 90 ry 0 rz 90 deg; joints [1.169, -72.71, 126.378, -178.55, 53.677, 179.141]
  MoveL 146 to (127.36, -41.26, 23.82) mm, rotated rx 90 ry 0 rz 90 deg; joints [1.226, -73.04, 126.846, -178.482, 53.816, 179.103]
  MoveL 147 to (121.15, -41.19, 22.72) mm, rotated rx 90 ry 0 rz 90 deg; joints [1.284, -73.373, 127.323, -178.412, 53.96, 179.065]
  MoveL 148 to (115.13, -41.16, 21.22) mm, rotated rx 90 ry 0 rz 90 deg; joints [1.363, -73.699, 127.783, -178.317, 54.095, 179.013]
  MoveL 149 to (109.45, -41.29, 18.9) mm, rotated rx 90 ry 0 rz 90 deg; joints [1.482, -74.014, 128.21, -178.173, 54.21, 178.931]
  MoveL 150 to (104.25, -41.31, 15.52) mm, rotated rx 90 ry 0 rz 90 deg; joints [1.654, -74.295, 128.598, -177.964, 54.32, 178.812]
  MoveL 151 to (99.57, -40.2, 11.27) mm, rotated rx 90 ry 0 rz 90 deg; joints [1.868, -74.486, 128.969, -177.706, 54.505, 178.667]
  MoveL 152 to (96.45, -38.41, 8.12) mm, rotated rx 90 ry 0 rz 90 deg; joints [2.027, -74.554, 129.236, -177.516, 54.707, 178.564]
  MoveL 153 to (93.71, -35.8, 5.55) mm, rotated rx 90 ry 0 rz 90 deg; joints [2.158, -74.557, 129.494, -177.364, 54.965, 178.486]
  MoveL 154 to (91.35, -32.35, 4.02) mm, rotated rx 90 ry 0 rz 90 deg; joints [2.238, -74.494, 129.742, -177.277, 55.278, 178.448]
  MoveL 155 to (89.22, -28.33, 3.44) mm, rotated rx 90 ry 0 rz 90 deg; joints [2.271, -74.386, 129.986, -177.249, 55.631, 178.446]
  MoveL 156 to (87.07, -24.08, 3.45) mm, rotated rx 90 ry 0 rz 90 deg; joints [2.274, -74.266, 130.237, -177.257, 56.002, 178.465]
  MoveL 157 to (84.65, -19.99, 3.7) mm, rotated rx 90 ry 0 rz 90 deg; joints [2.266, -74.167, 130.505, -177.278, 56.367, 178.491]
  MoveL 158 to (80.12, -14.75, 3.88) mm, rotated rx 90 ry 0 rz 90 deg; joints [2.267, -74.113, 130.954, -177.293, 56.87, 178.52]
  MoveL 159 to (74.83, -10.27, 3.79) mm, rotated rx 90 ry 0 rz 90 deg; joints [2.281, -74.138, 131.442, -177.29, 57.332, 178.536]
  MoveL 160 to (69.43, -5.9, 3.66) mm, rotated rx 90 ry 0 rz 90 deg; joints [2.299, -74.172, 131.934, -177.283, 57.791, 178.551]
  MoveL 161 to (64.56, -1, 3.71) mm, rotated rx 90 ry 0 rz 90 deg; joints [2.306, -74.141, 132.394, -177.288, 58.282, 178.574]
  Sollgeschwindigkeit (1000.0 mm/s)
  MoveL 162 to (64.56, -1, 3.71) mm, rotated rx 90 ry 0 rz 90 deg; joints [2.306, -74.141, 132.394, -177.288, 58.282, 178.574]
  MoveL 163 to (64.56, -1, 3.71) mm, rotated rx 90 ry 0 rz 90 deg; joints [2.306, -74.141, 132.394, -177.288, 58.282, 178.574]
  Sollgeschwindigkeit (1000.0 mm/s)
  MoveL 164 to (35.44, -1, 3.71) mm, rotated rx 90 ry 0 rz 90 deg; joints [2.367, -75.697, 134.575, -177.236, 58.907, 178.572]
  MoveL 165 to (35.44, -1, 3.71) mm, rotated rx 90 ry 0 rz 90 deg; joints [2.367, -75.697, 134.575, -177.236, 58.907, 178.572]
  MoveL 166 to (35.44, -1, 3.71) mm, rotated rx 90 ry 0 rz 90 deg; joints [2.367, -75.697, 134.575, -177.236, 58.907, 178.572]
  Sollgeschwindigkeit (50.0 mm/s)
  MoveL 167 to (30.57, -5.9, 3.66) mm, rotated rx 90 ry 0 rz 90 deg; joints [2.38, -76.263, 134.84, -177.212, 58.608, 178.547]
  MoveL 168 to (25.17, -10.27, 3.79) mm, rotated rx 90 ry 0 rz 90 deg; joints [2.384, -76.826, 135.153, -177.199, 58.357, 178.53]
  MoveL 169 to (19.88, -14.75, 3.88) mm, rotated rx 90 ry 0 rz 90 deg; joints [2.391, -77.393, 135.451, -177.182, 58.089, 178.51]
  MoveL 170 to (15.35, -19.99, 3.7) mm, rotated rx 90 ry 0 rz 90 deg; joints [2.411, -77.967, 135.673, -177.149, 57.739, 178.477]
  MoveL 171 to (12.93, -24.08, 3.45) mm, rotated rx 90 ry 0 rz 90 deg; joints [2.429, -78.352, 135.761, -177.117, 57.442, 178.448]
  MoveL 172 to (10.78, -28.33, 3.44) mm, rotated rx 90 ry 0 rz 90 deg; joints [2.435, -78.732, 135.824, -177.1, 57.126, 178.425]
  MoveL 173 to (8.65, -32.35, 4.02) mm, rotated rx 90 ry 0 rz 90 deg; joints [2.409, -79.098, 135.891, -177.121, 56.826, 178.424]
  MoveL 174 to (6.29, -35.8, 5.55) mm, rotated rx 90 ry 0 rz 90 deg; joints [2.333, -79.445, 135.988, -177.205, 56.575, 178.459]
  MoveL 175 to (3.55, -38.41, 8.12) mm, rotated rx 90 ry 0 rz 90 deg; joints [2.202, -79.767, 136.134, -177.356, 56.396, 178.536]
  MoveL 176 to (0.43, -40.2, 11.27) mm, rotated rx 90 ry 0 rz 90 deg; joints [2.04, -80.061, 136.327, -177.547, 56.291, 178.638]
  MoveL 177 to (-4.25, -41.31, 15.52) mm, rotated rx 90 ry 0 rz 90 deg; joints [1.822, -80.408, 136.65, -177.809, 56.262, 178.783]
  MoveL 178 to (-9.45, -41.29, 18.9) mm, rotated rx 90 ry 0 rz 90 deg; joints [1.648, -80.715, 137.034, -178.02, 56.335, 178.902]
  MoveL 179 to (-15.13, -41.16, 21.22) mm, rotated rx 90 ry 0 rz 90 deg; joints [1.532, -81.042, 137.451, -178.162, 56.422, 178.983]
  MoveL 180 to (-21.16, -41.19, 22.72) mm, rotated rx 90 ry 0 rz 90 deg; joints [1.458, -81.4, 137.887, -178.251, 56.498, 179.034]
  MoveL 181 to (-27.36, -41.26, 23.82) mm, rotated rx 90 ry 0 rz 90 deg; joints [1.407, -81.772, 138.332, -178.314, 56.572, 179.071]
  MoveL 182 to (-33.44, -41.28, 24.88) mm, rotated rx 90 ry 0 rz 90 deg; joints [1.356, -82.135, 138.768, -178.376, 56.644, 179.107]
  MoveL 183 to (-39.36, -41.27, 26.34) mm, rotated rx 90 ry 0 rz 90 deg; joints [1.283, -82.488, 139.193, -178.465, 56.715, 179.157]
  MoveL 184 to (-44.93, -41.25, 28.57) mm, rotated rx 90 ry 0 rz 90 deg; joints [1.166, -82.822, 139.593, -178.606, 56.779, 179.236]
  MoveL 185 to (-50, -41.25, 31.96) mm, rotated rx 90 ry 0 rz 90 deg; joints [0.981, -83.131, 139.958, -178.828, 56.832, 179.359]
  Sollgeschwindigkeit (1000.0 mm/s)
  MoveL 186 to (-50, -41.25, 31.96) mm, rotated rx 90 ry 0 rz 90 deg; joints [0.981, -83.131, 139.958, -178.828, 56.832, 179.359]
  MoveL 187 to (-50, -41.25, 31.96) mm, rotated rx 90 ry 0 rz 90 deg; joints [0.981, -83.131, 139.958, -178.828, 56.832, 179.359]
  Sollgeschwindigkeit (1000.0 mm/s)
  MoveL 188 to (-50, -40.49, 11.17) mm, rotated rx 90 ry 0 rz 90 deg; joints [2.147, -83.048, 139.936, -177.438, 56.914, 178.601]
  MoveL 189 to (-50, -40.49, 11.17) mm, rotated rx 90 ry 0 rz 90 deg; joints [2.147, -83.048, 139.936, -177.438, 56.914, 178.601]
  MoveL 190 to (-50, -40.49, 11.17) mm, rotated rx 90 ry 0 rz 90 deg; joints [2.147, -83.048, 139.936, -177.438, 56.914, 178.601]
  Sollgeschwindigkeit (50.0 mm/s)
  MoveL 191 to (-46.33, -40.39, 12.86) mm, rotated rx 90 ry 0 rz 90 deg; joints [2.045, -82.825, 139.683, -177.559, 56.881, 178.666]
  MoveL 192 to (-42.49, -40.49, 13.6) mm, rotated rx 90 ry 0 rz 90 deg; joints [1.996, -82.604, 139.409, -177.615, 56.828, 178.695]
  MoveL 193 to (-38.56, -40.66, 13.55) mm, rotated rx 90 ry 0 rz 90 deg; joints [1.991, -82.38, 139.125, -177.62, 56.768, 178.695]
  MoveL 194 to (-32.68, -40.73, 12.33) mm, rotated rx 90 ry 0 rz 90 deg; joints [2.047, -82.033, 138.701, -177.55, 56.692, 178.654]
  MoveL 195 to (-27.1, -40.17, 10.21) mm, rotated rx 90 ry 0 rz 90 deg; joints [2.152, -81.663, 138.31, -177.424, 56.673, 178.584]
  MoveL 196 to (-23.68, -39.22, 8.56) mm, rotated rx 90 ry 0 rz 90 deg; joints [2.236, -81.399, 138.083, -177.325, 56.713, 178.531]
  MoveL 197 to (-20.61, -37.64, 6.89) mm, rotated rx 90 ry 0 rz 90 deg; joints [2.32, -81.117, 137.896, -177.228, 56.809, 178.482]
  MoveL 198 to (-17.97, -35.32, 5.38) mm, rotated rx 90 ry 0 rz 90 deg; joints [2.396, -80.815, 137.756, -177.142, 56.974, 178.441]
  MoveL 199 to (-15.76, -32.33, 4.23) mm, rotated rx 90 ry 0 rz 90 deg; joints [2.453, -80.498, 137.663, -177.081, 57.199, 178.418]
  MoveL 200 to (-13.93, -28.93, 3.66) mm, rotated rx 90 ry 0 rz 90 deg; joints [2.48, -80.179, 137.608, -177.058, 57.464, 178.417]
  MoveL 201 to (-12.22, -25.42, 3.56) mm, rotated rx 90 ry 0 rz 90 deg; joints [2.481, -79.86, 137.564, -177.065, 57.738, 178.433]
  MoveL 202 to (-9.48, -21.06, 3.73) mm, rotated rx 90 ry 0 rz 90 deg; joints [2.465, -79.43, 137.463, -177.095, 58.066, 178.462]
  MoveL 203 to (-5.64, -17.69, 3.8) mm, rotated rx 90 ry 0 rz 90 deg; joints [2.453, -79, 137.258, -177.116, 58.29, 178.483]
  MoveL 204 to (-1.07, -15.06, 3.75) mm, rotated rx 90 ry 0 rz 90 deg; joints [2.445, -78.577, 136.981, -177.13, 58.436, 178.497]
  MoveL 205 to (3.61, -12.69, 3.72) mm, rotated rx 90 ry 0 rz 90 deg; joints [2.436, -78.167, 136.689, -177.144, 58.554, 178.509]
  MoveL 206 to (8.27, -10.42, 3.72) mm, rotated rx 90 ry 0 rz 90 deg; joints [2.426, -77.765, 136.395, -177.16, 58.661, 178.522]
  MoveL 207 to (17.27, -5.84, 3.76) mm, rotated rx 90 ry 0 rz 90 deg; joints [2.404, -76.984, 135.826, -177.192, 58.873, 178.547]
  MoveL 208 to (25.94, -0.5, 3.76) mm, rotated rx 90 ry 0 rz 90 deg; joints [2.385, -76.179, 135.29, -177.222, 59.141, 178.574]
  Sollgeschwindigkeit (1000.0 mm/s)
  MoveL 209 to (25.94, -0.5, 3.76) mm, rotated rx 90 ry 0 rz 90 deg; joints [2.385, -76.179, 135.29, -177.222, 59.141, 178.574]
  MoveL 210 to (25.94, -0.5, 3.76) mm, rotated rx 90 ry 0 rz 90 deg; joints [2.385, -76.179, 135.29, -177.222, 59.141, 178.574]
  Sollgeschwindigkeit (1000.0 mm/s)
  MoveL 211 to (74.06, -0.5, 3.76) mm, rotated rx 90 ry 0 rz 90 deg; joints [2.285, -73.608, 131.686, -177.309, 58.106, 178.577]
  MoveL 212 to (74.06, -0.5, 3.76) mm, rotated rx 90 ry 0 rz 90 deg; joints [2.285, -73.608, 131.686, -177.309, 58.106, 178.577]
  MoveL 213 to (74.06, -0.5, 3.76) mm, rotated rx 90 ry 0 rz 90 deg; joints [2.285, -73.608, 131.686, -177.309, 58.106, 178.577]
  Sollgeschwindigkeit (50.0 mm/s)
  MoveL 214 to (82.73, -5.84, 3.76) mm, rotated rx 90 ry 0 rz 90 deg; joints [2.267, -73.46, 130.928, -177.311, 57.496, 178.554]
  MoveL 215 to (91.73, -10.42, 3.72) mm, rotated rx 90 ry 0 rz 90 deg; joints [2.252, -73.244, 130.157, -177.313, 56.941, 178.533]
  MoveL 216 to (96.39, -12.69, 3.72) mm, rotated rx 90 ry 0 rz 90 deg; joints [2.243, -73.125, 129.758, -177.315, 56.661, 178.524]
  MoveL 217 to (101.07, -15.06, 3.75) mm, rotated rx 90 ry 0 rz 90 deg; joints [2.232, -73.008, 129.354, -177.319, 56.375, 178.514]
  MoveL 218 to (105.64, -17.69, 3.8) mm, rotated rx 90 ry 0 rz 90 deg; joints [2.221, -72.911, 128.953, -177.323, 56.071, 178.505]
  MoveL 219 to (109.48, -21.06, 3.73) mm, rotated rx 90 ry 0 rz 90 deg; joints [2.217, -72.892, 128.592, -177.316, 55.729, 178.488]
  MoveL 220 to (112.22, -25.42, 3.56) mm, rotated rx 90 ry 0 rz 90 deg; joints [2.221, -72.982, 128.294, -177.3, 55.342, 178.464]
  MoveL 221 to (113.93, -28.93, 3.66) mm, rotated rx 90 ry 0 rz 90 deg; joints [2.213, -73.08, 128.091, -177.3, 55.04, 178.452]
  MoveL 222 to (115.76, -32.33, 4.23) mm, rotated rx 90 ry 0 rz 90 deg; joints [2.182, -73.166, 127.882, -177.328, 54.745, 178.457]
  MoveL 223 to (117.97, -35.32, 5.38) mm, rotated rx 90 ry 0 rz 90 deg; joints [2.122, -73.208, 127.653, -177.392, 54.473, 178.484]
  MoveL 224 to (120.61, -37.64, 6.89) mm, rotated rx 90 ry 0 rz 90 deg; joints [2.045, -73.19, 127.405, -177.48, 54.241, 178.526]
  MoveL 225 to (123.68, -39.22, 8.56) mm, rotated rx 90 ry 0 rz 90 deg; joints [1.96, -73.109, 127.14, -177.579, 54.055, 178.578]
  MoveL 226 to (127.1, -40.17, 10.21) mm, rotated rx 90 ry 0 rz 90 deg; joints [1.876, -72.976, 126.861, -177.679, 53.907, 178.632]
  MoveL 227 to (132.68, -40.73, 12.33) mm, rotated rx 90 ry 0 rz 90 deg; joints [1.766, -72.705, 126.424, -177.81, 53.738, 178.704]
  MoveL 228 to (138.56, -40.66, 13.55) mm, rotated rx 90 ry 0 rz 90 deg; joints [1.7, -72.385, 125.974, -177.888, 53.608, 178.747]
  MoveL 229 to (142.49, -40.49, 13.6) mm, rotated rx 90 ry 0 rz 90 deg; joints [1.692, -72.163, 125.673, -177.896, 53.528, 178.749]
  MoveL 230 to (146.33, -40.39, 12.86) mm, rotated rx 90 ry 0 rz 90 deg; joints [1.721, -71.948, 125.375, -177.857, 53.446, 178.723]
  MoveL 231 to (150, -40.49, 11.17) mm, rotated rx 90 ry 0 rz 90 deg; joints [1.795, -71.752, 125.083, -177.762, 53.352, 178.664]
  Sollgeschwindigkeit (1000.0 mm/s)
  MoveL 232 to (150, -40.49, 11.17) mm, rotated rx 90 ry 0 rz 90 deg; joints [1.795, -71.752, 125.083, -177.762, 53.352, 178.664]
  MoveL 233 to (150, -40.49, 11.17) mm, rotated rx 90 ry 0 rz 90 deg; joints [1.795, -71.752, 125.083, -177.762, 53.352, 178.664]
  Sollgeschwindigkeit (1000.0 mm/s)
  MoveL 234 to (150, -28.4, 3.75) mm, rotated rx 90 ry 0 rz 90 deg; joints [2.143, -71.116, 125.312, -177.358, 54.225, 178.455]
  MoveL 235 to (150, -28.4, 3.75) mm, rotated rx 90 ry 0 rz 90 deg; joints [2.143, -71.116, 125.312, -177.358, 54.225, 178.455]
  MoveL 236 to (150, -28.4, 3.75) mm, rotated rx 90 ry 0 rz 90 deg; joints [2.143, -71.116, 125.312, -177.358, 54.225, 178.455]
  Sollgeschwindigkeit (50.0 mm/s)
  MoveL 237 to (146.28, -29.22, 3.75) mm, rotated rx 90 ry 0 rz 90 deg; joints [2.15, -71.357, 125.585, -177.351, 54.257, 178.452]
  MoveL 238 to (142.22, -28.97, 3.75) mm, rotated rx 90 ry 0 rz 90 deg; joints [2.157, -71.561, 125.907, -177.346, 54.374, 178.453]
  MoveL 239 to (138.31, -27.66, 3.75) mm, rotated rx 90 ry 0 rz 90 deg; joints [2.164, -71.703, 126.237, -177.344, 54.563, 178.459]
  MoveL 240 to (135.78, -26.02, 3.75) mm, rotated rx 90 ry 0 rz 90 deg; joints [2.168, -71.751, 126.466, -177.344, 54.744, 178.466]
  MoveL 241 to (133.82, -23.81, 3.75) mm, rotated rx 90 ry 0 rz 90 deg; joints [2.172, -71.738, 126.662, -177.347, 54.952, 178.476]
  MoveL 242 to (132.64, -21.07, 3.75) mm, rotated rx 90 ry 0 rz 90 deg; joints [2.174, -71.655, 126.807, -177.352, 55.181, 178.487]
  MoveL 243 to (132.33, -17.66, 3.75) mm, rotated rx 90 ry 0 rz 90 deg; joints [2.175, -71.488, 126.898, -177.359, 55.438, 178.501]
  MoveL 244 to (133.11, -14.37, 3.75) mm, rotated rx 90 ry 0 rz 90 deg; joints [2.173, -71.27, 126.901, -177.368, 55.659, 178.514]
  MoveL 245 to (134.92, -11.65, 3.75) mm, rotated rx 90 ry 0 rz 90 deg; joints [2.17, -71.027, 126.811, -177.377, 55.812, 178.525]
  MoveL 246 to (137.54, -9.53, 3.75) mm, rotated rx 90 ry 0 rz 90 deg; joints [2.165, -70.775, 126.648, -177.385, 55.9, 178.533]
  MoveL 247 to (141.76, -7.46, 3.75) mm, rotated rx 90 ry 0 rz 90 deg; joints [2.158, -70.442, 126.357, -177.395, 55.943, 178.541]
  MoveL 248 to (146.15, -6.05, 3.75) mm, rotated rx 90 ry 0 rz 90 deg; joints [2.15, -70.137, 126.04, -177.404, 55.931, 178.545]
  MoveL 249 to (150, -5.07, 3.75) mm, rotated rx 90 ry 0 rz 90 deg; joints [2.143, -69.884, 125.756, -177.412, 55.9, 178.548]
  Sollgeschwindigkeit (1000.0 mm/s)
  MoveL 250 to (150, -5.07, 3.75) mm, rotated rx 90 ry 0 rz 90 deg; joints [2.143, -69.884, 125.756, -177.412, 55.9, 178.548]
  MoveL 251 to (150, -5.07, 3.75) mm, rotated rx 90 ry 0 rz 90 deg; joints [2.143, -69.884, 125.756, -177.412, 55.9, 178.548]
  Sollgeschwindigkeit (1000.0 mm/s)
  MoveL 252 to (134.08, 0, 3.75) mm, rotated rx 90 ry 0 rz 90 deg; joints [2.171, -70.436, 127.09, -177.401, 56.681, 178.572]
  MoveL 253 to (134.08, 0, 3.75) mm, rotated rx 90 ry 0 rz 90 deg; joints [2.171, -70.436, 127.09, -177.401, 56.681, 178.572]
  MoveL 254 to (134.08, 0, 3.75) mm, rotated rx 90 ry 0 rz 90 deg; joints [2.171, -70.436, 127.09, -177.401, 56.681, 178.572]
  Sollgeschwindigkeit (50.0 mm/s)
  MoveL 255 to (133.99, -2.31, 3.75) mm, rotated rx 90 ry 0 rz 90 deg; joints [2.172, -70.567, 127.056, -177.396, 56.516, 178.563]
  MoveL 256 to (133.12, -4.45, 3.75) mm, rotated rx 90 ry 0 rz 90 deg; joints [2.173, -70.73, 127.085, -177.39, 56.382, 178.554]
  MoveL 257 to (131.64, -6.32, 3.75) mm, rotated rx 90 ry 0 rz 90 deg; joints [2.176, -70.91, 127.166, -177.384, 56.283, 178.547]
  MoveL 258 to (128.64, -8.39, 3.75) mm, rotated rx 90 ry 0 rz 90 deg; joints [2.181, -71.18, 127.36, -177.375, 56.207, 178.539]
  MoveL 259 to (125.24, -9.27, 3.75) mm, rotated rx 90 ry 0 rz 90 deg; joints [2.187, -71.408, 127.607, -177.368, 56.227, 178.536]
  MoveL 260 to (120.92, -8.94, 3.75) mm, rotated rx 90 ry 0 rz 90 deg; joints [2.195, -71.616, 127.947, -177.363, 56.358, 178.538]
  MoveL 261 to (116.63, -8.26, 3.75) mm, rotated rx 90 ry 0 rz 90 deg; joints [2.203, -71.805, 128.291, -177.358, 56.513, 178.542]
  MoveL 262 to (112.36, -7.56, 3.75) mm, rotated rx 90 ry 0 rz 90 deg; joints [2.211, -71.991, 128.632, -177.353, 56.669, 178.545]
  MoveL 263 to (102.41, -5.6, 3.75) mm, rotated rx 90 ry 0 rz 90 deg; joints [2.23, -72.405, 129.432, -177.343, 57.055, 178.554]
  MoveL 264 to (93.68, -3.23, 3.75) mm, rotated rx 90 ry 0 rz 90 deg; joints [2.247, -72.731, 130.144, -177.334, 57.441, 178.565]
  MoveL 265 to (85.1, 0, 3.75) mm, rotated rx 90 ry 0 rz 90 deg; joints [2.263, -72.996, 130.858, -177.328, 57.89, 178.579]
  Sollgeschwindigkeit (1000.0 mm/s)
  MoveL 266 to (85.1, 0, 3.75) mm, rotated rx 90 ry 0 rz 90 deg; joints [2.263, -72.996, 130.858, -177.328, 57.89, 178.579]
  MoveL 267 to (85.1, 0, 3.75) mm, rotated rx 90 ry 0 rz 90 deg; joints [2.263, -72.996, 130.858, -177.328, 57.89, 178.579]
  Sollgeschwindigkeit (1000.0 mm/s)
  MoveL 268 to (14.9, 0, 3.75) mm, rotated rx 90 ry 0 rz 90 deg; joints [2.409, -76.745, 136.117, -177.201, 59.401, 178.574]
  MoveL 269 to (14.9, 0, 3.75) mm, rotated rx 90 ry 0 rz 90 deg; joints [2.409, -76.745, 136.117, -177.201, 59.401, 178.574]
  MoveL 270 to (14.9, 0, 3.75) mm, rotated rx 90 ry 0 rz 90 deg; joints [2.409, -76.745, 136.117, -177.201, 59.401, 178.574]
  Sollgeschwindigkeit (50.0 mm/s)
  MoveL 271 to (6.32, -3.23, 3.75) mm, rotated rx 90 ry 0 rz 90 deg; joints [2.428, -77.419, 136.685, -177.175, 59.296, 178.557]
  MoveL 272 to (-2.41, -5.6, 3.75) mm, rotated rx 90 ry 0 rz 90 deg; joints [2.448, -78.05, 137.277, -177.151, 59.258, 178.543]
  MoveL 273 to (-12.36, -7.56, 3.75) mm, rotated rx 90 ry 0 rz 90 deg; joints [2.471, -78.729, 137.962, -177.125, 59.265, 178.53]
  MoveL 274 to (-16.63, -8.26, 3.75) mm, rotated rx 90 ry 0 rz 90 deg; joints [2.481, -79.013, 138.258, -177.113, 59.277, 178.524]
  MoveL 275 to (-20.92, -8.94, 3.75) mm, rotated rx 90 ry 0 rz 90 deg; joints [2.491, -79.298, 138.556, -177.102, 59.29, 178.519]
  MoveL 276 to (-25.24, -9.27, 3.75) mm, rotated rx 90 ry 0 rz 90 deg; joints [2.502, -79.563, 138.861, -177.091, 59.331, 178.515]
  MoveL 277 to (-28.64, -8.39, 3.75) mm, rotated rx 90 ry 0 rz 90 deg; joints [2.51, -79.697, 139.126, -177.086, 59.462, 178.518]
  MoveL 278 to (-31.64, -6.32, 3.75) mm, rotated rx 90 ry 0 rz 90 deg; joints [2.517, -79.729, 139.387, -177.084, 59.69, 178.528]
  MoveL 279 to (-33.12, -4.45, 3.75) mm, rotated rx 90 ry 0 rz 90 deg; joints [2.521, -79.688, 139.533, -177.086, 59.877, 178.536]
  MoveL 280 to (-33.99, -2.31, 3.75) mm, rotated rx 90 ry 0 rz 90 deg; joints [2.523, -79.594, 139.641, -177.089, 60.079, 178.547]
  MoveL 281 to (-34.08, 0, 3.75) mm, rotated rx 90 ry 0 rz 90 deg; joints [2.523, -79.444, 139.695, -177.095, 60.283, 178.559]
  Sollgeschwindigkeit (1000.0 mm/s)
  MoveL 282 to (-34.08, 0, 3.75) mm, rotated rx 90 ry 0 rz 90 deg; joints [2.523, -79.444, 139.695, -177.095, 60.283, 178.559]
  MoveL 283 to (-34.08, 0, 3.75) mm, rotated rx 90 ry 0 rz 90 deg; joints [2.523, -79.444, 139.695, -177.095, 60.283, 178.559]
  Sollgeschwindigkeit (1000.0 mm/s)
  MoveL 284 to (-50, -5.07, 3.75) mm, rotated rx 90 ry 0 rz 90 deg; joints [2.562, -80.687, 140.736, -177.044, 60.081, 178.524]
  MoveL 285 to (-50, -5.07, 3.75) mm, rotated rx 90 ry 0 rz 90 deg; joints [2.562, -80.687, 140.736, -177.044, 60.081, 178.524]
  MoveL 286 to (-50, -5.07, 3.75) mm, rotated rx 90 ry 0 rz 90 deg; joints [2.562, -80.687, 140.736, -177.044, 60.081, 178.524]
  Sollgeschwindigkeit (50.0 mm/s)
  MoveL 287 to (-46.15, -6.05, 3.75) mm, rotated rx 90 ry 0 rz 90 deg; joints [2.553, -80.534, 140.438, -177.05, 59.937, 178.521]
  MoveL 288 to (-41.76, -7.46, 3.75) mm, rotated rx 90 ry 0 rz 90 deg; joints [2.542, -80.379, 140.092, -177.057, 59.747, 178.516]
  MoveL 289 to (-37.54, -9.53, 3.75) mm, rotated rx 90 ry 0 rz 90 deg; joints [2.531, -80.277, 139.744, -177.062, 59.5, 178.508]
  MoveL 290 to (-34.92, -11.65, 3.75) mm, rotated rx 90 ry 0 rz 90 deg; joints [2.525, -80.269, 139.51, -177.062, 59.274, 178.498]
  MoveL 291 to (-33.11, -14.37, 3.75) mm, rotated rx 90 ry 0 rz 90 deg; joints [2.521, -80.345, 139.32, -177.059, 59.008, 178.485]
  MoveL 292 to (-32.33, -17.66, 3.75) mm, rotated rx 90 ry 0 rz 90 deg; joints [2.519, -80.515, 139.191, -177.052, 58.709, 178.468]
  MoveL 293 to (-32.64, -21.07, 3.75) mm, rotated rx 90 ry 0 rz 90 deg; joints [2.519, -80.755, 139.136, -177.042, 58.415, 178.45]
  MoveL 294 to (-33.82, -23.81, 3.75) mm, rotated rx 90 ry 0 rz 90 deg; joints [2.522, -81.001, 139.159, -177.032, 58.192, 178.434]
  MoveL 295 to (-35.78, -26.02, 3.75) mm, rotated rx 90 ry 0 rz 90 deg; joints [2.527, -81.257, 139.248, -177.021, 58.026, 178.421]
  MoveL 296 to (-38.31, -27.66, 3.75) mm, rotated rx 90 ry 0 rz 90 deg; joints [2.533, -81.511, 139.391, -177.01, 57.915, 178.411]
  MoveL 297 to (-42.22, -28.97, 3.75) mm, rotated rx 90 ry 0 rz 90 deg; joints [2.543, -81.825, 139.641, -176.996, 57.851, 178.401]
  MoveL 298 to (-46.28, -29.22, 3.75) mm, rotated rx 90 ry 0 rz 90 deg; joints [2.553, -82.081, 139.924, -176.985, 57.88, 178.396]
  MoveL 299 to (-50, -28.4, 3.75) mm, rotated rx 90 ry 0 rz 90 deg; joints [2.562, -82.246, 140.209, -176.978, 57.998, 178.398]
  Sollgeschwindigkeit (1000.0 mm/s)
  MoveL 300 to (-50, -28.4, 3.75) mm, rotated rx 90 ry 0 rz 90 deg; joints [2.562, -82.246, 140.209, -176.978, 57.998, 178.398]
  MoveL 301 to (-50, -28.4, 3.75) mm, rotated rx 90 ry 0 rz 90 deg; joints [2.562, -82.246, 140.209, -176.978, 57.998, 178.398]

--- program Pfad5 (robot KUKA KR 30 HA) ---
  Glatt(1)
  Sollgeschwindigkeit (1000.0 mm/s)
  Referenz erstellen.: Reference SW
  Werkzeug setzen: PlasticPos800
  Anzeigen PlasticPos800
  MoveJ 1 to (50, -38.85, 51.65) mm, rotated rx 90 ry 0 rz 90 deg; joints [-0.112, -77.197, 132.769, 179.865, 55.572, -179.923]
  MoveL 2 to (50, -38.85, 51.65) mm, rotated rx 90 ry 0 rz 90 deg; joints [-0.112, -77.197, 132.769, 179.865, 55.572, -179.923]
  MoveL 3 to (50, -38.85, 51.65) mm, rotated rx 90 ry 0 rz 90 deg; joints [-0.112, -77.197, 132.769, 179.865, 55.572, -179.923]
  MoveL 4 to (50, -38.85, 51.65) mm, rotated rx 90 ry 0 rz 90 deg; joints [-0.112, -77.197, 132.769, 179.865, 55.572, -179.923]
  Sollgeschwindigkeit (50.0 mm/s)
  MoveL 5 to (41.4, -38.88, 51.63) mm, rotated rx 90 ry 0 rz 90 deg; joints [-0.112, -77.683, 133.406, 179.865, 55.723, -179.924]
  MoveL 6 to (32.82, -39.2, 51.14) mm, rotated rx 90 ry 0 rz 90 deg; joints [-0.087, -78.186, 134.031, 179.895, 55.845, -179.941]
  MoveL 7 to (24.28, -39.97, 50.14) mm, rotated rx 90 ry 0 rz 90 deg; joints [-0.035, -78.716, 134.642, 179.957, 55.925, -179.976]
  MoveL 8 to (22, -40.34, 49.48) mm, rotated rx 90 ry 0 rz 90 deg; joints [-0.001, -78.868, 134.8, 179.999, 55.932, -180]
  MoveL 9 to (20.05, -40.65, 48.1) mm, rotated rx 90 ry 0 rz 90 deg; joints [0.071, -78.998, 134.936, 180.086, 55.937, -180.048]
  MoveL 10 to (18.53, -40.89, 46.07) mm, rotated rx 90 ry 0 rz 90 deg; joints [0.178, -79.1, 135.041, 180.215, 55.942, -180.121]
  MoveL 11 to (17.47, -41.07, 43.6) mm, rotated rx 90 ry 0 rz 90 deg; joints [0.308, -79.17, 135.114, 180.372, 55.945, -180.208]
  MoveL 12 to (16.87, -41.2, 40.01) mm, rotated rx 90 ry 0 rz 90 deg; joints [0.497, -79.211, 135.153, 180.6, 55.943, -180.336]
  MoveL 13 to (17.29, -41.25, 36.56) mm, rotated rx 90 ry 0 rz 90 deg; joints [0.679, -79.188, 135.118, 180.819, 55.933, -180.459]
  MoveL 14 to (18.81, -41.23, 33.72) mm, rotated rx 90 ry 0 rz 90 deg; joints [0.827, -79.097, 135.005, 180.999, 55.912, -180.56]
  MoveL 15 to (21.87, -41.2, 30.71) mm, rotated rx 90 ry 0 rz 90 deg; joints [0.982, -78.918, 134.778, 181.187, 55.866, -180.666]
  MoveL 16 to (24.9, -41.35, 27.7) mm, rotated rx 90 ry 0 rz 90 deg; joints [1.137, -78.75, 134.549, 181.375, 55.806, -180.773]
  MoveL 17 to (27.3, -41.63, 24.26) mm, rotated rx 90 ry 0 rz 90 deg; joints [1.314, -78.625, 134.36, 181.59, 55.745, -180.895]
  MoveL 18 to (29.82, -41.76, 19.45) mm, rotated rx 90 ry 0 rz 90 deg; joints [1.561, -78.483, 134.163, 181.89, 55.695, -181.065]
  MoveL 19 to (32.24, -41.12, 14.43) mm, rotated rx 90 ry 0 rz 90 deg; joints [1.818, -78.299, 133.989, 182.201, 55.71, -181.24]
  MoveL 20 to (34.88, -39.28, 9.61) mm, rotated rx 90 ry 0 rz 90 deg; joints [2.063, -78.034, 133.825, 182.494, 55.817, -181.402]
  MoveL 21 to (36.62, -37.37, 6.91) mm, rotated rx 90 ry 0 rz 90 deg; joints [2.199, -77.819, 133.733, 182.655, 55.943, -181.487]
  MoveL 22 to (38.19, -34.94, 4.93) mm, rotated rx 90 ry 0 rz 90 deg; joints [2.298, -77.584, 133.666, 182.768, 56.113, -181.544]
  MoveL 23 to (39.51, -32.01, 3.89) mm, rotated rx 90 ry 0 rz 90 deg; joints [2.349, -77.337, 133.63, 182.822, 56.325, -181.566]
  MoveL 24 to (40.8, -28.72, 3.61) mm, rotated rx 90 ry 0 rz 90 deg; joints [2.36, -77.072, 133.607, 182.829, 56.567, -181.559]
  MoveL 25 to (42.19, -25.66, 3.68) mm, rotated rx 90 ry 0 rz 90 deg; joints [2.354, -76.815, 133.57, 182.814, 56.786, -181.542]
  MoveL 26 to (44.08, -22.58, 3.79) mm, rotated rx 90 ry 0 rz 90 deg; joints [2.344, -76.529, 133.495, 182.796, 56.997, -181.524]
  MoveL 27 to (46.71, -19.51, 3.8) mm, rotated rx 90 ry 0 rz 90 deg; joints [2.338, -76.203, 133.364, 182.782, 57.192, -181.508]
  MoveL 28 to (48.43, -18.08, 3.78) mm, rotated rx 90 ry 0 rz 90 deg; joints [2.336, -76.024, 133.266, 182.777, 57.272, -181.502]
  MoveL 29 to (50, -17.29, 3.75) mm, rotated rx 90 ry 0 rz 90 deg; joints [2.334, -75.892, 133.165, 182.774, 57.304, -181.499]
  MoveL 30 to (50, -17.29, 3.75) mm, rotated rx 90 ry 0 rz 90 deg; joints [2.334, -75.892, 133.165, 182.774, 57.304, -181.499]
  MoveL 31 to (51.57, -18.08, 3.78) mm, rotated rx 90 ry 0 rz 90 deg; joints [2.329, -75.852, 133.031, 182.771, 57.21, -181.501]
  MoveL 32 to (53.29, -19.51, 3.8) mm, rotated rx 90 ry 0 rz 90 deg; joints [2.324, -75.843, 132.874, 182.77, 57.062, -181.507]
  MoveL 33 to (55.92, -22.58, 3.79) mm, rotated rx 90 ry 0 rz 90 deg; joints [2.32, -75.879, 132.613, 182.774, 56.766, -181.521]
  MoveL 34 to (57.81, -25.66, 3.68) mm, rotated rx 90 ry 0 rz 90 deg; joints [2.321, -75.953, 132.407, 182.784, 56.484, -181.538]
  MoveL 35 to (59.2, -28.72, 3.61) mm, rotated rx 90 ry 0 rz 90 deg; joints [2.322, -76.053, 132.237, 182.794, 56.216, -181.555]
  MoveL 36 to (60.49, -32.01, 3.89) mm, rotated rx 90 ry 0 rz 90 deg; joints [2.305, -76.171, 132.071, 182.783, 55.931, -181.56]
  MoveL 37 to (61.81, -34.94, 4.93) mm, rotated rx 90 ry 0 rz 90 deg; joints [2.25, -76.267, 131.911, 182.725, 55.675, -181.537]
  MoveL 38 to (63.38, -37.37, 6.91) mm, rotated rx 90 ry 0 rz 90 deg; joints [2.147, -76.321, 131.746, 182.607, 55.453, -181.479]
  MoveL 39 to (65.12, -39.28, 9.61) mm, rotated rx 90 ry 0 rz 90 deg; joints [2.008, -76.337, 131.58, 182.443, 55.268, -181.393]
  MoveL 40 to (67.76, -41.12, 14.43) mm, rotated rx 90 ry 0 rz 90 deg; joints [1.761, -76.302, 131.354, 182.149, 55.071, -181.231]
  MoveL 41 to (70.18, -41.76, 19.45) mm, rotated rx 90 ry 0 rz 90 deg; joints [1.506, -76.211, 131.169, 181.839, 54.972, -181.056]
  MoveL 42 to (72.7, -41.63, 24.26) mm, rotated rx 90 ry 0 rz 90 deg; joints [1.262, -76.069, 130.992, 181.542, 54.932, -180.886]
  MoveL 43 to (75.1, -41.35, 27.7) mm, rotated rx 90 ry 0 rz 90 deg; joints [1.087, -75.924, 130.823, 181.329, 54.906, -180.764]
  MoveL 44 to (78.13, -41.2, 30.71) mm, rotated rx 90 ry 0 rz 90 deg; joints [0.934, -75.751, 130.603, 181.143, 54.857, -180.658]
  MoveL 45 to (81.19, -41.23, 33.72) mm, rotated rx 90 ry 0 rz 90 deg; joints [0.782, -75.585, 130.376, 180.958, 54.794, -180.552]
  MoveL 46 to (82.71, -41.25, 36.56) mm, rotated rx 90 ry 0 rz 90 deg; joints [0.64, -75.504, 130.263, 180.784, 54.762, -180.452]
  MoveL 47 to (83.13, -41.2, 40.01) mm, rotated rx 90 ry 0 rz 90 deg; joints [0.469, -75.48, 130.235, 180.574, 54.757, -180.331]
  MoveL 48 to (82.53, -41.07, 43.6) mm, rotated rx 90 ry 0 rz 90 deg; joints [0.291, -75.507, 130.285, 180.356, 54.779, -180.205]
  MoveL 49 to (81.47, -40.89, 46.07) mm, rotated rx 90 ry 0 rz 90 deg; joints [0.169, -75.556, 130.369, 180.206, 54.813, -180.119]
  MoveL 50 to (79.95, -40.65, 48.1) mm, rotated rx 90 ry 0 rz 90 deg; joints [0.068, -75.628, 130.49, 180.083, 54.862, -180.048]
  MoveL 51 to (78, -40.34, 49.48) mm, rotated rx 90 ry 0 rz 90 deg; joints [-0.001, -75.719, 130.644, 179.999, 54.925, -180]
  MoveL 52 to (75.72, -39.97, 50.14) mm, rotated rx 90 ry 0 rz 90 deg; joints [-0.034, -75.825, 130.823, 179.959, 54.999, -179.976]
  MoveL 53 to (67.18, -39.2, 51.14) mm, rotated rx 90 ry 0 rz 90 deg; joints [-0.084, -76.257, 131.481, 179.897, 55.224, -179.941]
  MoveL 54 to (58.6, -38.88, 51.63) mm, rotated rx 90 ry 0 rz 90 deg; joints [-0.11, -76.717, 132.128, 179.866, 55.411, -179.924]
  MoveL 55 to (50, -38.85, 51.65) mm, rotated rx 90 ry 0 rz 90 deg; joints [-0.112, -77.197, 132.769, 179.865, 55.572, -179.923]
  Sollgeschwindigkeit (1000.0 mm/s)
  MoveL 56 to (50, -38.85, 51.65) mm, rotated rx 90 ry 0 rz 90 deg; joints [-0.112, -77.197, 132.769, 179.865, 55.572, -179.923]
  MoveL 57 to (50, -38.85, 51.65) mm, rotated rx 90 ry 0 rz 90 deg; joints [-0.112, -77.197, 132.769, 179.865, 55.572, -179.923]
  Sollgeschwindigkeit (1000.0 mm/s)
  MoveL 58 to (50, -41.25, 44.41) mm, rotated rx 90 ry 0 rz 90 deg; joints [0.258, -77.334, 132.714, 180.314, 55.381, -180.178]
  MoveL 59 to (50, -41.25, 44.41) mm, rotated rx 90 ry 0 rz 90 deg; joints [0.258, -77.334, 132.714, 180.314, 55.381, -180.178]
  MoveL 60 to (50, -41.25, 44.41) mm, rotated rx 90 ry 0 rz 90 deg; joints [0.258, -77.334, 132.714, 180.314, 55.381, -180.178]
  Sollgeschwindigkeit (50.0 mm/s)
  MoveL 61 to (45.62, -41.25, 43.91) mm, rotated rx 90 ry 0 rz 90 deg; joints [0.285, -77.58, 133.039, 180.346, 55.459, -180.196]
  MoveL 62 to (41.42, -41.25, 43.16) mm, rotated rx 90 ry 0 rz 90 deg; joints [0.325, -77.817, 133.349, 180.394, 55.532, -180.223]
  MoveL 63 to (38.6, -41.25, 42.58) mm, rotated rx 90 ry 0 rz 90 deg; joints [0.355, -77.977, 133.557, 180.43, 55.581, -180.243]
  MoveL 64 to (35.9, -41.25, 41.66) mm, rotated rx 90 ry 0 rz 90 deg; joints [0.404, -78.13, 133.756, 180.489, 55.627, -180.276]
  MoveL 65 to (34.18, -41.25, 39.31) mm, rotated rx 90 ry 0 rz 90 deg; joints [0.526, -78.226, 133.881, 180.637, 55.657, -180.36]
  MoveL 66 to (33.35, -41.24, 35.37) mm, rotated rx 90 ry 0 rz 90 deg; joints [0.731, -78.27, 133.939, 180.885, 55.672, -180.499]
  MoveL 67 to (33.65, -41.22, 31.56) mm, rotated rx 90 ry 0 rz 90 deg; joints [0.928, -78.249, 133.913, 181.124, 55.67, -180.634]
  MoveL 68 to (34.41, -41.27, 27.86) mm, rotated rx 90 ry 0 rz 90 deg; joints [1.119, -78.205, 133.851, 181.355, 55.654, -180.765]
  MoveL 69 to (35.45, -41.41, 23.18) mm, rotated rx 90 ry 0 rz 90 deg; joints [1.36, -78.148, 133.764, 181.648, 55.627, -180.931]
  MoveL 70 to (36.64, -41.36, 18.45) mm, rotated rx 90 ry 0 rz 90 deg; joints [1.603, -78.071, 133.669, 181.943, 55.613, -181.098]
  MoveL 71 to (38.13, -40.8, 13.62) mm, rotated rx 90 ry 0 rz 90 deg; joints [1.85, -77.946, 133.561, 182.241, 55.636, -181.266]
  MoveL 72 to (39.64, -39.56, 9.61) mm, rotated rx 90 ry 0 rz 90 deg; joints [2.054, -77.781, 133.468, 182.486, 55.712, -181.401]
  MoveL 73 to (41.11, -37.31, 6.47) mm, rotated rx 90 ry 0 rz 90 deg; joints [2.213, -77.562, 133.402, 182.673, 55.869, -181.501]
  MoveL 74 to (42.58, -33.91, 4.58) mm, rotated rx 90 ry 0 rz 90 deg; joints [2.307, -77.277, 133.363, 182.779, 56.117, -181.55]
  MoveL 75 to (44.02, -30.73, 3.87) mm, rotated rx 90 ry 0 rz 90 deg; joints [2.34, -77.011, 133.324, 182.812, 56.346, -181.559]
  MoveL 76 to (45.95, -27.27, 3.65) mm, rotated rx 90 ry 0 rz 90 deg; joints [2.347, -76.701, 133.256, 182.813, 56.587, -181.55]
  MoveL 77 to (47.84, -24.64, 3.68) mm, rotated rx 90 ry 0 rz 90 deg; joints [2.342, -76.443, 133.172, 182.8, 56.76, -181.536]
  MoveL 78 to (48.85, -23.61, 3.72) mm, rotated rx 90 ry 0 rz 90 deg; joints [2.338, -76.327, 133.119, 182.793, 56.823, -181.529]
  MoveL 79 to (50, -22.99, 3.75) mm, rotated rx 90 ry 0 rz 90 deg; joints [2.334, -76.227, 133.046, 182.788, 56.85, -181.525]
  MoveL 80 to (50, -22.99, 3.75) mm, rotated rx 90 ry 0 rz 90 deg; joints [2.334, -76.227, 133.046, 182.788, 56.85, -181.525]
  MoveL 81 to (51.15, -23.61, 3.72) mm, rotated rx 90 ry 0 rz 90 deg; joints [2.333, -76.2, 132.947, 182.789, 56.778, -181.529]
  MoveL 82 to (52.16, -24.64, 3.68) mm, rotated rx 90 ry 0 rz 90 deg; joints [2.333, -76.205, 132.85, 182.792, 56.676, -181.535]
  MoveL 83 to (54.05, -27.27, 3.65) mm, rotated rx 90 ry 0 rz 90 deg; joints [2.331, -76.253, 132.653, 182.797, 56.431, -181.548]
  MoveL 84 to (55.98, -30.73, 3.87) mm, rotated rx 90 ry 0 rz 90 deg; joints [2.315, -76.347, 132.435, 182.789, 56.12, -181.556]
  MoveL 85 to (57.42, -33.91, 4.58) mm, rotated rx 90 ry 0 rz 90 deg; joints [2.277, -76.451, 132.261, 182.752, 55.841, -181.546]
  MoveL 86 to (58.89, -37.31, 6.47) mm, rotated rx 90 ry 0 rz 90 deg; joints [2.178, -76.566, 132.081, 182.641, 55.543, -181.495]
  MoveL 87 to (60.36, -39.56, 9.61) mm, rotated rx 90 ry 0 rz 90 deg; joints [2.016, -76.618, 131.93, 182.452, 55.336, -181.395]
  MoveL 88 to (61.87, -40.8, 13.62) mm, rotated rx 90 ry 0 rz 90 deg; joints [1.811, -76.611, 131.799, 182.206, 55.208, -181.259]
  MoveL 89 to (63.36, -41.36, 18.45) mm, rotated rx 90 ry 0 rz 90 deg; joints [1.565, -76.567, 131.686, 181.908, 55.133, -181.091]
  MoveL 90 to (64.55, -41.41, 23.18) mm, rotated rx 90 ry 0 rz 90 deg; joints [1.325, -76.51, 131.605, 181.616, 55.105, -180.925]
  MoveL 91 to (65.59, -41.27, 27.86) mm, rotated rx 90 ry 0 rz 90 deg; joints [1.088, -76.45, 131.538, 181.327, 55.095, -180.76]
  MoveL 92 to (66.35, -41.22, 31.56) mm, rotated rx 90 ry 0 rz 90 deg; joints [0.901, -76.409, 131.487, 181.099, 55.083, -180.629]
  MoveL 93 to (66.65, -41.24, 35.37) mm, rotated rx 90 ry 0 rz 90 deg; joints [0.709, -76.396, 131.468, 180.865, 55.076, -180.495]
  MoveL 94 to (65.82, -41.25, 39.31) mm, rotated rx 90 ry 0 rz 90 deg; joints [0.512, -76.445, 131.533, 180.624, 55.089, -180.357]
  MoveL 95 to (64.1, -41.25, 41.66) mm, rotated rx 90 ry 0 rz 90 deg; joints [0.394, -76.542, 131.663, 180.48, 55.122, -180.274]
  MoveL 96 to (61.4, -41.25, 42.58) mm, rotated rx 90 ry 0 rz 90 deg; joints [0.348, -76.693, 131.865, 180.424, 55.172, -180.242]
  MoveL 97 to (58.58, -41.25, 43.16) mm, rotated rx 90 ry 0 rz 90 deg; joints [0.32, -76.851, 132.075, 180.389, 55.225, -180.222]
  MoveL 98 to (54.38, -41.25, 43.91) mm, rotated rx 90 ry 0 rz 90 deg; joints [0.283, -77.087, 132.388, 180.344, 55.302, -180.196]
  MoveL 99 to (50, -41.25, 44.41) mm, rotated rx 90 ry 0 rz 90 deg; joints [0.258, -77.334, 132.714, 180.314, 55.381, -180.178]
  Sollgeschwindigkeit (1000.0 mm/s)
  MoveL 100 to (50, -41.25, 44.41) mm, rotated rx 90 ry 0 rz 90 deg; joints [0.258, -77.334, 132.714, 180.314, 55.381, -180.178]
  MoveL 101 to (50, -41.25, 44.41) mm, rotated rx 90 ry 0 rz 90 deg; joints [0.258, -77.334, 132.714, 180.314, 55.381, -180.178]
  Sollgeschwindigkeit (1000.0 mm/s)
  MoveL 102 to (50, -41.25, 34.01) mm, rotated rx 90 ry 0 rz 90 deg; joints [0.789, -77.328, 132.707, 180.959, 55.382, -180.545]
  MoveL 103 to (50, -41.25, 34.01) mm, rotated rx 90 ry 0 rz 90 deg; joints [0.789, -77.328, 132.707, 180.959, 55.382, -180.545]
  MoveL 104 to (50, -41.25, 34.01) mm, rotated rx 90 ry 0 rz 90 deg; joints [0.789, -77.328, 132.707, 180.959, 55.382, -180.545]
  Sollgeschwindigkeit (50.0 mm/s)
  MoveL 105 to (47.54, -41.17, 33.12) mm, rotated rx 90 ry 0 rz 90 deg; joints [0.837, -77.462, 132.89, 181.016, 55.432, -180.577]
  MoveL 106 to (45.56, -41.21, 31.05) mm, rotated rx 90 ry 0 rz 90 deg; joints [0.944, -77.574, 133.034, 181.146, 55.466, -180.65]
  MoveL 107 to (44.02, -41.28, 28.52) mm, rotated rx 90 ry 0 rz 90 deg; joints [1.075, -77.662, 133.143, 181.305, 55.488, -180.74]
  MoveL 108 to (42.9, -41.35, 25.95) mm, rotated rx 90 ry 0 rz 90 deg; joints [1.209, -77.726, 133.22, 181.467, 55.503, -180.831]
  MoveL 109 to (41.78, -41.35, 20.71) mm, rotated rx 90 ry 0 rz 90 deg; joints [1.479, -77.783, 133.294, 181.795, 55.524, -181.016]
  MoveL 110 to (41.91, -41.03, 15.28) mm, rotated rx 90 ry 0 rz 90 deg; joints [1.758, -77.748, 133.28, 182.133, 55.551, -181.207]
  MoveL 111 to (42.51, -40.36, 11.73) mm, rotated rx 90 ry 0 rz 90 deg; joints [1.94, -77.67, 133.243, 182.351, 55.596, -181.329]
  MoveL 112 to (43.34, -39.01, 8.54) mm, rotated rx 90 ry 0 rz 90 deg; joints [2.102, -77.538, 133.204, 182.545, 55.692, -181.435]
  MoveL 113 to (44.38, -36.75, 5.98) mm, rotated rx 90 ry 0 rz 90 deg; joints [2.231, -77.345, 133.171, 182.696, 55.856, -181.514]
  MoveL 114 to (45.3, -34.77, 4.8) mm, rotated rx 90 ry 0 rz 90 deg; joints [2.29, -77.176, 133.144, 182.763, 55.998, -181.546]
  MoveL 115 to (46.5, -32.46, 4.09) mm, rotated rx 90 ry 0 rz 90 deg; joints [2.324, -76.974, 133.104, 182.798, 56.161, -181.559]
  MoveL 116 to (48.06, -29.92, 3.77) mm, rotated rx 90 ry 0 rz 90 deg; joints [2.337, -76.739, 133.042, 182.808, 56.335, -181.558]
  MoveL 117 to (49.06, -28.63, 3.73) mm, rotated rx 90 ry 0 rz 90 deg; joints [2.337, -76.608, 132.995, 182.806, 56.419, -181.553]
  MoveL 118 to (50, -27.82, 3.75) mm, rotated rx 90 ry 0 rz 90 deg; joints [2.334, -76.509, 132.943, 182.8, 56.466, -181.548]
  MoveL 119 to (50, -27.82, 3.75) mm, rotated rx 90 ry 0 rz 90 deg; joints [2.334, -76.509, 132.943, 182.8, 56.466, -181.548]
  MoveL 120 to (50.94, -28.63, 3.73) mm, rotated rx 90 ry 0 rz 90 deg; joints [2.333, -76.504, 132.856, 182.802, 56.383, -181.552]
  MoveL 121 to (51.94, -29.92, 3.77) mm, rotated rx 90 ry 0 rz 90 deg; joints [2.329, -76.523, 132.753, 182.801, 56.262, -181.557]
  MoveL 122 to (53.5, -32.46, 4.09) mm, rotated rx 90 ry 0 rz 90 deg; joints [2.309, -76.584, 132.583, 182.785, 56.03, -181.557]
  MoveL 123 to (54.7, -34.77, 4.8) mm, rotated rx 90 ry 0 rz 90 deg; joints [2.271, -76.651, 132.444, 182.745, 55.824, -181.543]
  MoveL 124 to (55.62, -36.75, 5.98) mm, rotated rx 90 ry 0 rz 90 deg; joints [2.209, -76.716, 132.335, 182.676, 55.649, -181.511]
  MoveL 125 to (56.66, -39.01, 8.54) mm, rotated rx 90 ry 0 rz 90 deg; joints [2.078, -76.792, 132.215, 182.523, 55.45, -181.431]
  MoveL 126 to (57.49, -40.36, 11.73) mm, rotated rx 90 ry 0 rz 90 deg; joints [1.914, -76.828, 132.131, 182.328, 55.325, -181.325]
  MoveL 127 to (58.09, -41.03, 15.28) mm, rotated rx 90 ry 0 rz 90 deg; joints [1.733, -76.838, 132.08, 182.109, 55.259, -181.202]
  MoveL 128 to (58.22, -41.35, 20.71) mm, rotated rx 90 ry 0 rz 90 deg; joints [1.458, -76.858, 132.074, 181.775, 55.229, -181.012]
  MoveL 129 to (57.1, -41.35, 25.95) mm, rotated rx 90 ry 0 rz 90 deg; joints [1.193, -76.927, 132.166, 181.453, 55.248, -180.828]
  MoveL 130 to (55.98, -41.28, 28.52) mm, rotated rx 90 ry 0 rz 90 deg; joints [1.064, -76.989, 132.255, 181.295, 55.273, -180.738]
  MoveL 131 to (54.44, -41.21, 31.05) mm, rotated rx 90 ry 0 rz 90 deg; joints [0.937, -77.074, 132.374, 181.14, 55.306, -180.649]
  MoveL 132 to (52.46, -41.17, 33.12) mm, rotated rx 90 ry 0 rz 90 deg; joints [0.833, -77.185, 132.525, 181.013, 55.344, -180.576]
  MoveL 133 to (50, -41.25, 34.01) mm, rotated rx 90 ry 0 rz 90 deg; joints [0.789, -77.328, 132.707, 180.959, 55.382, -180.545]
  Sollgeschwindigkeit (1000.0 mm/s)
  MoveL 134 to (50, -41.25, 34.01) mm, rotated rx 90 ry 0 rz 90 deg; joints [0.789, -77.328, 132.707, 180.959, 55.382, -180.545]
  MoveL 135 to (50, -41.25, 34.01) mm, rotated rx 90 ry 0 rz 90 deg; joints [0.789, -77.328, 132.707, 180.959, 55.382, -180.545]

--- program Pfad6 (robot KUKA KR 30 HA) ---
  Glatt(1)
  Sollgeschwindigkeit (1000.0 mm/s)
  Referenz erstellen.: Reference SW
  Werkzeug setzen: PlasticPos800
  Anzeigen PlasticPos800
  MoveJ 1 to (20.69, 0, 56.25) mm, rotated rx 90 ry 0 rz 90 deg; joints [-0.356, -76.483, 135.759, 179.586, 59.277, -179.788]
  MoveL 2 to (20.69, 0, 56.25) mm, rotated rx 90 ry 0 rz 90 deg; joints [-0.356, -76.483, 135.759, 179.586, 59.277, -179.788]
  MoveL 3 to (20.69, 0, 56.25) mm, rotated rx 90 ry 0 rz 90 deg; joints [-0.356, -76.483, 135.759, 179.586, 59.277, -179.788]
  MoveL 4 to (20.69, 0, 56.25) mm, rotated rx 90 ry 0 rz 90 deg; joints [-0.356, -76.483, 135.759, 179.586, 59.277, -179.788]
  Sollgeschwindigkeit (50.0 mm/s)
  MoveL 5 to (22.63, -4.6, 56.24) mm, rotated rx 90 ry 0 rz 90 deg; joints [-0.355, -76.665, 135.524, 179.586, 58.86, -179.786]
  MoveL 6 to (25.24, -8.42, 56.25) mm, rotated rx 90 ry 0 rz 90 deg; joints [-0.355, -76.759, 135.254, 179.584, 58.495, -179.783]
  MoveL 7 to (28.4, -11.75, 56.28) mm, rotated rx 90 ry 0 rz 90 deg; joints [-0.355, -76.791, 134.953, 179.582, 58.162, -179.779]
  MoveL 8 to (31.96, -14.9, 56.29) mm, rotated rx 90 ry 0 rz 90 deg; joints [-0.355, -76.787, 134.624, 179.581, 57.838, -179.777]
  MoveL 9 to (34.49, -17.04, 56.28) mm, rotated rx 90 ry 0 rz 90 deg; joints [-0.353, -76.777, 134.392, 179.582, 57.615, -179.776]
  MoveL 10 to (37.11, -19.32, 56.25) mm, rotated rx 90 ry 0 rz 90 deg; joints [-0.351, -76.77, 134.15, 179.584, 57.38, -179.776]
  MoveL 11 to (39.78, -21.76, 56.19) mm, rotated rx 90 ry 0 rz 90 deg; joints [-0.347, -76.768, 133.9, 179.587, 57.132, -179.776]
  MoveL 12 to (42.51, -24.11, 56.14) mm, rotated rx 90 ry 0 rz 90 deg; joints [-0.343, -76.757, 133.648, 179.59, 56.891, -179.776]
  MoveL 13 to (45.72, -25.96, 56.1) mm, rotated rx 90 ry 0 rz 90 deg; joints [-0.34, -76.688, 133.37, 179.593, 56.682, -179.776]
  MoveL 14 to (50, -26.64, 56.09) mm, rotated rx 90 ry 0 rz 90 deg; joints [-0.338, -76.491, 133.036, 179.594, 56.546, -179.776]
  MoveL 15 to (54.28, -25.96, 56.1) mm, rotated rx 90 ry 0 rz 90 deg; joints [-0.338, -76.215, 132.732, 179.595, 56.518, -179.777]
  MoveL 16 to (57.49, -24.11, 56.14) mm, rotated rx 90 ry 0 rz 90 deg; joints [-0.339, -75.931, 132.531, 179.594, 56.601, -179.777]
  MoveL 17 to (60.22, -21.76, 56.19) mm, rotated rx 90 ry 0 rz 90 deg; joints [-0.341, -75.645, 132.376, 179.593, 56.732, -179.777]
  MoveL 18 to (62.89, -19.32, 56.25) mm, rotated rx 90 ry 0 rz 90 deg; joints [-0.343, -75.357, 132.227, 179.591, 56.87, -179.776]
  MoveL 19 to (65.51, -17.04, 56.28) mm, rotated rx 90 ry 0 rz 90 deg; joints [-0.344, -75.082, 132.077, 179.59, 56.995, -179.777]
  MoveL 20 to (68.04, -14.9, 56.29) mm, rotated rx 90 ry 0 rz 90 deg; joints [-0.343, -74.82, 131.929, 179.591, 57.109, -179.778]
  MoveL 21 to (71.6, -11.75, 56.28) mm, rotated rx 90 ry 0 rz 90 deg; joints [-0.342, -74.445, 131.723, 179.594, 57.279, -179.78]
  MoveL 22 to (74.76, -8.42, 56.25) mm, rotated rx 90 ry 0 rz 90 deg; joints [-0.339, -74.082, 131.55, 179.597, 57.469, -179.783]
  MoveL 23 to (77.37, -4.6, 56.24) mm, rotated rx 90 ry 0 rz 90 deg; joints [-0.338, -73.72, 131.426, 179.6, 57.706, -179.787]
  MoveL 24 to (79.31, 0, 56.25) mm, rotated rx 90 ry 0 rz 90 deg; joints [-0.338, -73.348, 131.365, 179.602, 58.017, -179.789]
  Sollgeschwindigkeit (1000.0 mm/s)
  MoveL 25 to (79.31, 0, 56.25) mm, rotated rx 90 ry 0 rz 90 deg; joints [-0.338, -73.348, 131.365, 179.602, 58.017, -179.789]
  MoveL 26 to (79.31, 0, 56.25) mm, rotated rx 90 ry 0 rz 90 deg; joints [-0.338, -73.348, 131.365, 179.602, 58.017, -179.789]

